(* IEC 61131-3 sources: plcassist-cli/packages/volt-lsp-iec/test-corpus/pro2193/Device/Plc Logic/Application/09 Misc/Library Manager/AlarmManager (part 2) *)

(* ---- ACK_ALARMSTATEMACHINE.fb ---- *)
FUNCTION_BLOCK ACK_ALARMSTATEMACHINE
END_FUNCTION_BLOCK

METHOD DOACKNOWLEDGE : AlarmState
VAR_INPUT
	ECURRENTSTATE : AlarmState;
END_VAR
VAR_OUTPUT
	ESTATETRANSITION : AlarmStateTransition;
END_VAR
END_METHOD

METHOD DOACTIVATE : AlarmState
VAR_INPUT
	ECURRENTSTATE : AlarmState;
END_VAR
END_METHOD

METHOD DODEACTIVATE : AlarmState
VAR_INPUT
	ECURRENTSTATE : AlarmState;
END_VAR
VAR_OUTPUT
	ESTATETRANSITION : AlarmStateTransition;
END_VAR
END_METHOD

(* ---- ACK_ALARMSTATEMACHINE_NOCONFIRM.fb ---- *)
FUNCTION_BLOCK ACK_ALARMSTATEMACHINE_NOCONFIRM EXTENDS Ack_AlarmStateMachine
END_FUNCTION_BLOCK

METHOD DOACKNOWLEDGE : AlarmState
VAR_INPUT
	ECURRENTSTATE : AlarmState;
END_VAR
VAR_OUTPUT
	ESTATETRANSITION : AlarmStateTransition;
END_VAR
END_METHOD

(* ---- ACK_REP_ACK_ALARMSTATEMACHINE.fb ---- *)
FUNCTION_BLOCK ACK_REP_ACK_ALARMSTATEMACHINE
END_FUNCTION_BLOCK

METHOD DOACKNOWLEDGE : AlarmState
VAR_INPUT
	ECURRENTSTATE : AlarmState;
END_VAR
VAR_OUTPUT
	ESTATETRANSITION : AlarmStateTransition;
END_VAR
END_METHOD

METHOD DOACTIVATE : AlarmState
VAR_INPUT
	ECURRENTSTATE : AlarmState;
END_VAR
END_METHOD

METHOD DODEACTIVATE : AlarmState
VAR_INPUT
	ECURRENTSTATE : AlarmState;
END_VAR
VAR_OUTPUT
	ESTATETRANSITION : AlarmStateTransition;
END_VAR
END_METHOD

(* ---- ACK_REP_ACK_ALARMSTATEMACHINE_NOCONFIRM.fb ---- *)
FUNCTION_BLOCK ACK_REP_ACK_ALARMSTATEMACHINE_NOCONFIRM EXTENDS Ack_Rep_Ack_AlarmStateMachine
END_FUNCTION_BLOCK

METHOD DOACKNOWLEDGE : AlarmState
VAR_INPUT
	ECURRENTSTATE : AlarmState;
END_VAR
VAR_OUTPUT
	ESTATETRANSITION : AlarmStateTransition;
END_VAR
END_METHOD

METHOD DODEACTIVATE : AlarmState
VAR_INPUT
	ECURRENTSTATE : AlarmState;
END_VAR
VAR_OUTPUT
	ESTATETRANSITION : AlarmStateTransition;
END_VAR
END_METHOD

(* ---- ACK_REP_ALARMSTATEMACHINE.fb ---- *)
FUNCTION_BLOCK ACK_REP_ALARMSTATEMACHINE
END_FUNCTION_BLOCK

METHOD DOACKNOWLEDGE : AlarmState
VAR_INPUT
	ECURRENTSTATE : AlarmState;
END_VAR
VAR_OUTPUT
	ESTATETRANSITION : AlarmStateTransition;
END_VAR
END_METHOD

METHOD DOACTIVATE : AlarmState
VAR_INPUT
	ECURRENTSTATE : AlarmState;
END_VAR
END_METHOD

METHOD DODEACTIVATE : AlarmState
VAR_INPUT
	ECURRENTSTATE : AlarmState;
END_VAR
VAR_OUTPUT
	ESTATETRANSITION : AlarmStateTransition;
END_VAR
END_METHOD

(* ---- ACK_REP_ALARMSTATEMACHINE_NOCONFIRM.fb ---- *)
FUNCTION_BLOCK ACK_REP_ALARMSTATEMACHINE_NOCONFIRM EXTENDS Ack_Rep_AlarmStateMachine
END_FUNCTION_BLOCK

METHOD DOACKNOWLEDGE : AlarmState
VAR_INPUT
	ECURRENTSTATE : AlarmState;
END_VAR
VAR_OUTPUT
	ESTATETRANSITION : AlarmStateTransition;
END_VAR
END_METHOD

METHOD DODEACTIVATE : AlarmState
VAR_INPUT
	ECURRENTSTATE : AlarmState;
END_VAR
VAR_OUTPUT
	ESTATETRANSITION : AlarmStateTransition;
END_VAR
END_METHOD

(* ---- ACTIVEALARMSTEMPSTORAGE.fb ---- *)
FUNCTION_BLOCK ACTIVEALARMSTEMPSTORAGE
VAR
	_LSTALARMSINFO : COL.IDoubleLinkedList := NULL;
	_LINKEDLISTFACTORY : COL.LinkedListFactory;
	_LISTVALUEELEMFACTORY : ListElementFactory;
END_VAR
END_FUNCTION_BLOCK

METHOD RESTOREALARMS : BOOL
END_METHOD

METHOD STOREALARMS : COL.COLLECTION_ERROR
VAR_INPUT
	PALARMGROUP : IAlarmGroup6;
END_VAR
END_METHOD

METHOD PRVRESTOREADDITIONALALARMINFO : INT
VAR_INPUT
	ITFLISTELEMENT : IListElement;
	PALARMUSED : POINTER TO Alarm;
END_VAR
END_METHOD

METHOD PRVSETALARMINFO : INT
VAR_INPUT
	PALARMSTORED : POINTER TO Alarm;
	PALARMUSED : POINTER TO Alarm;
	ITFLISTELEMENT : IListElement;
END_VAR
END_METHOD

METHOD PRVSTOREACTIVEALARM : BOOL
VAR_INPUT
	ITFLISTELEMENT : IListElement;
	PALARM : POINTER TO Alarm;
END_VAR
END_METHOD

METHOD PRVSTOREALARMS : BOOL
VAR_INPUT
	PALARMGROUP : IAlarmGroup6;
END_VAR
END_METHOD

(* ---- ADAPTERDATABLOCK.fb ---- *)
FUNCTION_BLOCK ADAPTERDATABLOCK
VAR_INPUT
	M_PARRITFALARMSFROMHISTORY : POINTER TO ARRAY [0..0] OF IAlarm2;
	M_PARRALARMSGRPFORHISTORY : POINTER TO ARRAY [0..10] OF POINTER TO AlarmGroupAdapter;
	M_PARRALARMSCLFORHISTORY : POINTER TO ARRAY [0..10] OF POINTER TO AlarmClassAdapter;
	M_ICOUNTALARMSFROMHISTORY : INT;
	M_PAITFALARMCONFIGURATIONS : POINTER TO ARRAY [0..0] OF IAlarmConfiguration;
	M_ICOUNTCONFIGURATIONS : INT;
	M_DITOTALCOUNTROWS : DINT;
END_VAR
VAR
	M_ALARMADAPTER : AlarmAdapter;
	M_ICOUNTROWS : INT;
END_VAR
END_FUNCTION_BLOCK

METHOD GETALARMMETAOBJECTSTUB : IAlarmMetaObjectStub3
VAR_INPUT
	IROW : INT;
	IOFFSET : INT;
END_VAR
END_METHOD

METHOD GETCOUNTROWS : INT
END_METHOD

METHOD HASALARMS : BOOL
END_METHOD

METHOD SETCOUNTROWS : BOOL
VAR_INPUT
	ICOUNT : INT;
END_VAR
END_METHOD

METHOD SETTOTALCOUNTROWS : BOOL
VAR_INPUT
	DICOUNT : DINT;
END_VAR
END_METHOD

(* ---- ALARM.fb ---- *)
FUNCTION_BLOCK ALARM
VAR_INPUT
	M_UIID : ALARM_ID;
	M_UDIID : UDINT;
	M_PALATCHVARIABLES : POINTER TO ARRAY [0..255] OF POINTER TO ValueTypeBundle;
	M_USICOUNTLATCHVARIABLES : USINT;
	M_XDYNVARIABLES : BOOL;
	M_PAPLACEHOLDERINFO : POINTER TO ARRAY [0..255] OF POINTER TO PlaceholderInfo;
	M_USICOUNTMESSAGES : USINT;
END_VAR
VAR
	M_ITFALARMOBSERVATIONTYPE : IAlarmObservationType;
	M_ITFDEACTIVATOR : IDeactivator;
	M_ITFALARMCLASS : IAlarmClass;
	M_ITFALARMGROUP : IAlarmGroup;
	M_ITFALARMGROUPTEMPLATE : IAlarmGroup;
	M_TONDELAYTIME : TIME;
	M_TOFFDELAYTIME : TIME;
	M_LITIMESTAMPACTIVE : Timestamp;
	M_LITIMESTAMPINACTIVE : Timestamp;
	M_LITIMESTAMPACKNOWLEDGE : Timestamp;
	M_LITIMESTAMPLAST : Timestamp;
	M_LITIMESTAMPONDELAY : Timestamp;
	M_LITIMESTAMPOFFDELAY : Timestamp;
	M_IOFFSETACTIVE : INT := -1;
	M_IOFFSETINACTIVE : INT := -1;
	M_IOFFSETACKNOWLEDGE : INT := -1;
	M_IOFFSETLAST : INT := -1;
	M_ESTATE : AlarmState;
	M_XTOACKNOWLEDGE : BOOL;
	M_TIGGERVALUE : ValueTypeBundle;
	M_CURRENTVALUE : ValueTypeBundle;
	M_ITFHIGHERPRIOALARM : IAlarm;
	M_ROWID : CAA.IDENT;
	M_XADDTOLISTOFACTIVEALARMS : BOOL;
	M_XCYCLICUPDATE : BOOL;
	M_XISDEACTIVATEDPREV : BOOL;
	M_SREMDEVICENAME : STRING;
	M_CMTACTIVE : AlarmComment;
	M_CMTACTIVEACK : AlarmComment;
	M_CMTWAITINGCONF : AlarmComment;
	M_CMTNORMAL : AlarmComment;
	M_UDIREALARMREPEATCOUNT : UDINT;
	M_USICOUNTLATCHVARIABLESORIGINAL : INT := -1;
	M_ITFALARM : IAlarm := THIS^;
	ACKNOWLEDGE : BOOL;
	ADDTOLISTOFACTIVEALARMS : BOOL;
	ALARMGROUPTEMPLATE : IAlarmGroup;
	COMMENTACTIVE : POINTER TO WSTRING;
	COMMENTACTIVEACK : POINTER TO WSTRING;
	COMMENTNORMAL : POINTER TO WSTRING;
	COMMENTWAITINGCONF : POINTER TO WSTRING;
	COUNTLATCHVARIABLESORIGINAL : INT;
	CYCLICUPDATE : BOOL;
	ISDEACTIVATEDPREV : BOOL;
	KINDOF : EAlarmType;
	OFFSETACKNOWLEDGE : INT;
	OFFSETACTIVE : INT;
	OFFSETINACTIVE : INT;
	OFFSETLAST : INT;
	REALARMREPEATCOUNT : UDINT;
	REMOTEDEVICENAME : STRING;
	USERIDCOMMENTACTIVE : POINTER TO WSTRING;
	USERIDCOMMENTACTIVEACK : POINTER TO WSTRING;
	USERIDCOMMENTNORMAL : POINTER TO WSTRING;
	USERIDCOMMENTWAITINGCONF : POINTER TO WSTRING;
END_VAR
END_FUNCTION_BLOCK

METHOD ANALYZEPLACEHOLDERS3 : BOOL
VAR_INPUT
	STRINGTYPE : __SYSTEM.TYPE_CLASS;
	IWHICHMESSAGE : INT;
END_VAR
END_METHOD

METHOD FB_EXIT : BOOL
VAR_INPUT
	BINCOPYCODE : BOOL;
END_VAR
END_METHOD

METHOD GETALARMCLASS : IAlarmClass
END_METHOD

METHOD GETALARMGROUP : IAlarmGroup
END_METHOD

METHOD GETHIGHERPRIOALARM : IAlarm
END_METHOD

METHOD GETID : ALARM_ID
END_METHOD

METHOD GETINTERNALID : UDINT
END_METHOD

METHOD GETMESSAGE : CharBufferPtr
VAR_INPUT
	STRINGTYPE : __SYSTEM.TYPE_CLASS;
END_VAR
END_METHOD

METHOD GETOBSERVATIONTYPE : IAlarmObservationType
END_METHOD

METHOD GETROWID : CAA.IDENT
END_METHOD

METHOD GETSTATE : AlarmState
END_METHOD

METHOD ISDEACTIVATED : BOOL
END_METHOD

METHOD SETALARMCLASS
VAR_INPUT
	ITFALARMCLASS : IAlarmClass;
END_VAR
END_METHOD

METHOD SETALARMGROUP
VAR_INPUT
	ITFALARMGROUP : IAlarmGroup;
END_VAR
END_METHOD

METHOD SETHIGHERPRIOALARM
VAR_INPUT
	ITFALARM : IAlarm;
END_VAR
END_METHOD

METHOD SETOBSERVATIONTYPE
VAR_INPUT
	ITFOBSERVATIONTYPE : IAlarmObservationType;
END_VAR
END_METHOD

METHOD SETROWID
VAR_INPUT
	ROWID : CAA.IDENT;
END_VAR
END_METHOD

METHOD SETTIMESTAMP
VAR_INPUT
	LICURRTIMESTAMP : Timestamp;
	ESTATE : AlarmState;
	ESTATETRANSITION : AlarmStateTransition;
END_VAR
END_METHOD

METHOD SETALARMSTATE
VAR_INPUT
	EALARMSTATE : AlarmState;
END_VAR
END_METHOD

METHOD SETCURRENTVALUE
VAR_INPUT
	ITFTYPEDVALUECURRENT : ITypedValue;
END_VAR
END_METHOD

METHOD SETID
VAR_INPUT
	UIID : ALARM_ID;
END_VAR
END_METHOD

METHOD SETINTERNALID
VAR_INPUT
	UDIID : UDINT;
END_VAR
END_METHOD

METHOD SETLATCHVAR1VALUE
VAR_INPUT
	ITFTYPEDVALUELATCHVAR1 : ITypedValue;
END_VAR
END_METHOD

METHOD SETLATCHVAR2VALUE
VAR_INPUT
	ITFTYPEDVALUELATCHVAR2 : ITypedValue;
END_VAR
END_METHOD

METHOD SETTIMESTAMPACKNOWLEDGE
VAR_INPUT
	LITIMESTAMPACKNOWLEDGE : Timestamp;
END_VAR
END_METHOD

METHOD SETTIMESTAMPACTIVE
VAR_INPUT
	LITIMESTAMPACTIVE : Timestamp;
END_VAR
END_METHOD

METHOD SETTIMESTAMPINACTIVE
VAR_INPUT
	LITIMESTAMPINACTIVE : Timestamp;
END_VAR
END_METHOD

METHOD SETTIMESTAMPLAST
VAR_INPUT
	LITIMESTAMPLAST : Timestamp;
END_VAR
END_METHOD

METHOD SETTRIGGERVALUE
VAR_INPUT
	ITFTYPEDVALUETRIGGER : ITypedValue;
END_VAR
END_METHOD

METHOD GETCOUNTLATCHVARIABLES : USINT
END_METHOD

METHOD GETCOUNTMESSAGES : USINT
END_METHOD

METHOD GETLATCHVARVALUE : ITypedValue
VAR_INPUT
	IWHICHLATCHVAR : INT;
END_VAR
END_METHOD

METHOD GETMESSAGE2 : CharBufferPtr
VAR_INPUT
	STRINGTYPE : __SYSTEM.TYPE_CLASS;
	IWHICHMESSAGE : INT;
END_VAR
END_METHOD

METHOD SETLATCHVARVALUE
VAR_INPUT
	IWHICHLATCHVAR : INT;
	ITFTYPEDVALUELATCHVAR : ITypedValue;
END_VAR
END_METHOD

METHOD SETTIMESTAMP2
VAR_INPUT
	LICURRTIMESTAMP : Timestamp;
	IOFFSET : INT;
	ESTATE : AlarmState;
	ESTATETRANSITION : AlarmStateTransition;
END_VAR
END_METHOD

METHOD GETLATCHVARIABLESADDRESS
VAR_OUTPUT
	PALATCHVARIABLES : POINTER TO BYTE;
	USICOUNTLATCHVARIABLES : USINT;
END_VAR
END_METHOD

METHOD SETLATCHVARIABLESADDRESS
VAR_INPUT
	PALATCHVARIABLES : POINTER TO BYTE;
	USICOUNTLATCHVARIABLES : USINT;
END_VAR
END_METHOD

METHOD ANALYZEPLACEHOLDERS
VAR_INPUT
	STRINGTYPE : __SYSTEM.TYPE_CLASS;
END_VAR
END_METHOD

METHOD GETCOUNTPLACEHOLDERS : SINT
END_METHOD

METHOD GETPLACEHOLDER : PlaceholderOccurrence
VAR_INPUT
	SIWHICHPLACEHOLDER : SINT;
END_VAR
END_METHOD

METHOD HASPLACEHOLDERREQUIRINGCYCLICALLYUPDATE : BOOL
END_METHOD

METHOD HASPLACEHOLDERS : BOOL
END_METHOD

METHOD ISOPTIMIZEDPLACEHOLDERREPLACEMENTSUPPORTED : BOOL
END_METHOD

METHOD ANALYZEPLACEHOLDERS2
VAR_INPUT
	STRINGTYPE : __SYSTEM.TYPE_CLASS;
	IWHICHMESSAGE : INT;
END_VAR
END_METHOD

METHOD GETCOUNTPLACEHOLDERS2 : SINT
VAR_INPUT
	IWHICHMESSAGE : INT;
END_VAR
END_METHOD

METHOD GETPLACEHOLDER2 : PlaceholderOccurrence
VAR_INPUT
	SIWHICHPLACEHOLDER : SINT;
	IWHICHMESSAGE : INT;
END_VAR
END_METHOD

METHOD HASPLACEHOLDERREQUIRINGCYCLICALLYUPDATE2 : BOOL
VAR_INPUT
	IWHICHMESSAGE : INT;
END_VAR
END_METHOD

METHOD HASPLACEHOLDERS2 : BOOL
VAR_INPUT
	IWHICHMESSAGE : INT;
END_VAR
END_METHOD

METHOD ISOPTIMIZEDPLACEHOLDERREPLACEMENTSUPPORTED2 : BOOL
VAR_INPUT
	IWHICHMESSAGE : INT;
END_VAR
END_METHOD

METHOD CANBEACTIVATED : BOOL
END_METHOD

METHOD CANBEDEACTIVATED : BOOL
END_METHOD

METHOD DETERMINETIMESTAMP
VAR_INPUT
	ESTATE : AlarmState;
	ESTATETRANSITION : AlarmStateTransition;
END_VAR
END_METHOD

METHOD GETALARM : IAlarm
END_METHOD

METHOD GETLATCHVARIABLESADDRESSDIRECT : BOOL
VAR_OUTPUT
	PALATCHVARIABLES : POINTER TO BYTE;
	USICOUNTLATCHVARIABLES : USINT;
END_VAR
END_METHOD

METHOD HANDLEAUTORESETDIGITALALARMS : BOOL
END_METHOD

METHOD INVALIDATEMESSAGEFLAGS
END_METHOD

METHOD RETRIEVECURRENTVALUE
VAR_INPUT
	ITFVALUEPROVIDER : IValueProvider;
END_VAR
END_METHOD

METHOD RETRIEVELATCHVARVALUE
VAR_INPUT
	IWHICHLATCHVARIABLE : INT;
	ITFVALUEPROVIDER : IValueProvider;
END_VAR
END_METHOD

METHOD RETRIEVELATCHVARVALUES
VAR_INPUT
	ITFVALUEPROVIDER : IValueProvider;
END_VAR
END_METHOD

METHOD RETRIEVETRIGGERVALUE
VAR_INPUT
	ITFVALUEPROVIDER : IValueProvider;
END_VAR
END_METHOD

METHOD SETACKNOWLEDGE : BOOL
VAR_INPUT
	PWSCOMMENT : POINTER TO WSTRING;
	PWSUSERID : POINTER TO WSTRING;
END_VAR
END_METHOD

METHOD SETACKNOWLEDGELOCKED : BOOL
VAR_INPUT
	PWSCOMMENT : POINTER TO WSTRING;
	PWSUSERID : POINTER TO WSTRING;
END_VAR
END_METHOD

METHOD SETCOMMENT : UDINT
VAR_INPUT
	PWSCOMMENT : POINTER TO WSTRING;
	PWSUSERID : POINTER TO WSTRING;
END_VAR
END_METHOD

METHOD SETCOMMENTDIRECTLY
VAR_INPUT
	PALARMOTHER : POINTER TO Alarm;
END_VAR
END_METHOD

METHOD SETDEACTIVATOR
VAR_INPUT
	ITFDEACTIVATOR : IDeactivator;
END_VAR
END_METHOD

METHOD SETOFFDELAYTIME
VAR_INPUT
	TTIME : TIME;
END_VAR
END_METHOD

METHOD SETONDELAYTIME
VAR_INPUT
	TTIME : TIME;
END_VAR
END_METHOD

METHOD SETREALARMREPEATCOUNTDIRECTLY
VAR_INPUT
	UDIREALARMREPEATCOUNT : UDINT;
END_VAR
END_METHOD

METHOD SETSTATE
VAR_INPUT
	ESTATE : AlarmState;
	ESTATETRANSITION : AlarmStateTransition;
END_VAR
END_METHOD

METHOD SETTIMESTAMPOFFDELAY
VAR_INPUT
	XRESET : BOOL;
END_VAR
END_METHOD

METHOD SETTIMESTAMPDELAY
VAR_INPUT
	XRESET : BOOL;
	TDELAY : TIME;
END_VAR
VAR_IN_OUT
	LITIMESTAMPDELAY : Timestamp;
END_VAR
END_METHOD

METHOD SETTIMESTAMPOFFDELAYDIRECTLY
VAR_INPUT
	LITIMESTAMPOFFDELAY : Timestamp;
END_VAR
END_METHOD

METHOD SETTIMESTAMPONDELAY
VAR_INPUT
	XRESET : BOOL;
END_VAR
END_METHOD

METHOD SETTIMESTAMPONDELAYDIRECTLY
VAR_INPUT
	LITIMESTAMPONDELAY : Timestamp;
END_VAR
END_METHOD

METHOD SETTRIGGERVALUEDIRECTLY
VAR_INPUT
	TRIGGERVALUE : ValueTypeBundle;
END_VAR
END_METHOD

METHOD ISCOMMENTTOSTATENORMAL : BOOL
END_METHOD

METHOD RESETALARMCOMMENTS
END_METHOD

METHOD RESETFORNEWCYCLE
END_METHOD

METHOD PRVCHECKPOSTALARM
VAR_INPUT
	ESTATE : AlarmState;
	EOLDSTATE : AlarmState;
	XFORCEUPDATE : BOOL;
END_VAR
END_METHOD

METHOD PRVCOPYFROMTYPEDVALUE
VAR_INPUT
	PVALUETYPEBUNDLETARGET : POINTER TO ValueTypeBundle;
	ITFTYPEDVALUESOURCE : ITypedValue;
END_VAR
END_METHOD

METHOD GETTIMESTAMPACKNOWLEDGE : Timestamp
END_METHOD

METHOD GETTIMESTAMPACTIVE : Timestamp
END_METHOD

METHOD GETTIMESTAMPINACTIVE : Timestamp
END_METHOD

METHOD GETTIMESTAMPLAST : Timestamp
END_METHOD

METHOD GETCURRENTVALUE : ITypedValue
END_METHOD

METHOD GETLATCHVAR1VALUE : ITypedValue
END_METHOD

METHOD GETLATCHVAR2VALUE : ITypedValue
END_METHOD

METHOD GETTRIGGERVALUE : ITypedValue
END_METHOD

(* ---- ALARMADAPTER.fb ---- *)
FUNCTION_BLOCK ALARMADAPTER
VAR_INPUT
	M_ITFALARM2 : IAlarm2;
	M_PALARMGROUP : POINTER TO AlarmGroupAdapter;
	M_PALARMCLASS : POINTER TO AlarmClassAdapter;
	M_PAITFALARMCONFIGURATIONS : POINTER TO ARRAY [0..0] OF IAlarmConfiguration;
	M_ICOUNTCONFIGURATIONS : INT;
END_VAR
VAR
	M_PLIVALUE : POINTER TO LINT;
	ALARMCLASSINTERNALID : UDINT;
	ALARMGROUPINTERNALID : UDINT;
	ALARMINTERNALID : UDINT;
	OFFSETACKNOWLEDGE : INT;
	OFFSETACTIVE : INT;
	OFFSETINACTIVE : INT;
	OFFSETLAST : INT;
	PROXYNAME : STRING;
	REMOTEALARMCLASSNAME : STRING;
	REMOTEALARMGROUPNAME : STRING;
	REMOTEALARMSTRINGID : STRING;
	REMOTEALARMTEXTLIST : STRING;
END_VAR
END_FUNCTION_BLOCK

METHOD INITIALIZE
END_METHOD

METHOD SETALARM
VAR_INPUT
	PALARM : POINTER TO Alarm;
END_VAR
END_METHOD

METHOD SETALARMGROUP
VAR_INPUT
	SALARMGROUP : STRING;
END_VAR
END_METHOD

METHOD SETCURRENTVALUE
VAR_INPUT
	ITFTYPEDVALUECURRENT : AlarmManager_Interfaces.ITypedValue;
END_VAR
END_METHOD

METHOD SETID
VAR_INPUT
	UIID : ALARM_ID;
END_VAR
END_METHOD

METHOD SETLATCHVAR1VALUE
VAR_INPUT
	ITFTYPEDVALUELATCHVAR1 : AlarmManager_Interfaces.ITypedValue;
END_VAR
END_METHOD

METHOD SETLATCHVAR2VALUE
VAR_INPUT
	ITFTYPEDVALUELATCHVAR2 : AlarmManager_Interfaces.ITypedValue;
END_VAR
END_METHOD

METHOD SETSTATE
VAR_INPUT
	ISTATE : INT;
END_VAR
END_METHOD

METHOD SETTIMESTAMPACKNOWLEDGE
VAR_INPUT
	LITIMESTAMPACKNOWLEDGE : Timestamp;
END_VAR
END_METHOD

METHOD SETTIMESTAMPACTIVE
VAR_INPUT
	LITIMESTAMPACTIVE : Timestamp;
END_VAR
END_METHOD

METHOD SETTIMESTAMPINACTIVE
VAR_INPUT
	LITIMESTAMPINACTIVE : Timestamp;
END_VAR
END_METHOD

METHOD SETTIMESTAMPLAST
VAR_INPUT
	LITIMESTAMPLAST : Timestamp;
END_VAR
END_METHOD

METHOD SETTRIGGERVALUE
VAR_INPUT
	ITFTYPEDVALUETRIGGER : AlarmManager_Interfaces.ITypedValue;
END_VAR
END_METHOD

METHOD GETPRIORITY : BYTE
END_METHOD

METHOD SETPRIORITY
VAR_INPUT
	BYPRIORITY : BYTE;
END_VAR
END_METHOD

METHOD GETCOUNTLATCHVARIABLES : USINT
END_METHOD

METHOD SETLATCHVARVALUE
VAR_INPUT
	IWHICHLATCHVAR : INT;
	ITFTYPEDVALUELATCHVAR : ITypedValue;
END_VAR
END_METHOD

METHOD PRVPREPARELATCHVARVALUE : ValueTypeBundle
VAR_INPUT
	ITFTYPEDVALUELATCHVAR : AlarmManager_Interfaces.ITypedValue;
END_VAR
END_METHOD

METHOD GETALARM : POINTER TO Alarm
END_METHOD

METHOD GETALARMGROUP : STRING
END_METHOD

METHOD GETCHECKSUM : UDINT
END_METHOD

METHOD GETCURRENTVALUE : AlarmManager_Interfaces.ITypedValue
END_METHOD

METHOD GETID : ALARM_ID
END_METHOD

METHOD GETLATCHVAR1VALUE : AlarmManager_Interfaces.ITypedValue
END_METHOD

METHOD GETLATCHVAR2VALUE : AlarmManager_Interfaces.ITypedValue
END_METHOD

METHOD GETSTATE : INT
END_METHOD

METHOD GETTIMESTAMPACKNOWLEDGE : Timestamp
END_METHOD

METHOD GETTIMESTAMPACTIVE : Timestamp
END_METHOD

METHOD GETTIMESTAMPINACTIVE : Timestamp
END_METHOD

METHOD GETTIMESTAMPLAST : Timestamp
END_METHOD

METHOD GETTRIGGERVALUE : AlarmManager_Interfaces.ITypedValue
END_METHOD

METHOD SETACKNOWLEDGE
VAR_INPUT
	BACKNOWLEDGEMULTIPLE : BOOL;
END_VAR
END_METHOD

METHOD SWAPVALUES
END_METHOD

METHOD GETACKNOWLEDGE : BOOL
END_METHOD

METHOD GETACKNOWLEDGEMULTIPLE : BOOL
END_METHOD

METHOD GETALARMCLASS : STRING
END_METHOD

METHOD GETSTRINGID : STRING
END_METHOD

METHOD GETTESTLISTNAME : STRING
END_METHOD

METHOD RESETACKNOWLEDGE
END_METHOD

METHOD SETALARMCLASS
VAR_INPUT
	SALARMCLASS : STRING;
END_VAR
END_METHOD

METHOD SETSTRINGID
VAR_INPUT
	SID : STRING;
END_VAR
END_METHOD

METHOD SETTESTLISTNAME
VAR_INPUT
	STESTLISTNAME : STRING;
END_VAR
END_METHOD

METHOD SETACKNOWLEDGE2
VAR_INPUT
	BACKNOWLEDGEMULTIPLE : BOOL;
END_VAR
END_METHOD

METHOD GETLATCHVARVALUE : ITypedValue2
VAR_INPUT
	IWHICHLATCHVAR : INT;
END_VAR
END_METHOD

(* ---- ALARMAPIOBSERVATIONTYPE.fb ---- *)
FUNCTION_BLOCK ALARMAPIOBSERVATIONTYPE
VAR
	M_XISACTIVE : BOOL;
	ALARMCONDITIONACTIVE : BOOL;
END_VAR
END_FUNCTION_BLOCK

METHOD ISACTIVE : BOOL
VAR_INPUT
	ECURRSTATE : AlarmState;
END_VAR
END_METHOD

METHOD ISIMMEDIATELYACTIVE : BOOL
END_METHOD

(* ---- ALARMCLASS.fb ---- *)
FUNCTION_BLOCK ALARMCLASS
VAR
	M_UDIID : UDINT;
	M_USIPRIORITY : USINT;
	M_XARCHIVING : BOOL;
	M_EACKNOWLEDGEMETHOD : AcknowledgeMethod;
	M_XACKNOWLEDGESEPARATELY : BOOL;
	M_XAUTORESETDIGITALALARMS : BOOL;
	M_XACKINSTEADOFCONFIRM : BOOL;
	M_PAITFALARMNOTIFIABLES : POINTER TO ARRAY [0..0] OF IAlarmNotifiable;
	M_ICOUNTNOTIFIABLES : INT;
	M_SNAME : STRING;
	M_PAPDISPLAYOPTIONS : POINTER TO ARRAY [AlarmState.Normal..AlarmState.ActiveAcknowledged] OF POINTER TO DisplayOptions;
	M_TREALARMTIME : TIME;
	REALARMTIME : TIME;
END_VAR
END_FUNCTION_BLOCK

METHOD SETACKINSTEADOFCONFIRM : BOOL
VAR_INPUT
	XACKINSTEADOFCONFIRM : BOOL;
END_VAR
END_METHOD

METHOD SETACKNOWLEDGEMETHOD
VAR_INPUT
	EACKNOWLEDGEMETHOD : AcknowledgeMethod;
END_VAR
END_METHOD

METHOD SETACKNOWLEDGESEPARATELY
VAR_INPUT
	XACKNOWLEDGESEPARATELY : BOOL;
END_VAR
END_METHOD

METHOD SETALARMNOTIFIABLES
END_METHOD

METHOD SETARCHIVING
VAR_INPUT
	XARCHIVING : BOOL;
END_VAR
END_METHOD

METHOD SETAUTORESETDIGITALALARMS
VAR_INPUT
	XAUTORESETDIGITALALARMS : BOOL;
END_VAR
END_METHOD

METHOD SETDISPLAYOPTIONS
END_METHOD

METHOD SETINTERNALID
VAR_INPUT
	UDIID : UDINT;
END_VAR
END_METHOD

METHOD SETNAME
VAR_INPUT
	SNAME : STRING;
END_VAR
END_METHOD

METHOD SETPRIORITY
VAR_INPUT
	USIPRIORITY : USINT;
END_VAR
END_METHOD

METHOD SETREALARMTIME
VAR_INPUT
	T : TIME;
END_VAR
END_METHOD

METHOD GETACKNOWLEDGEMETHOD : AcknowledgeMethod
END_METHOD

METHOD GETALARMSTATEMACHINE : IAlarmStateMachine
END_METHOD

METHOD GETDISPLAYOPTIONS : POINTER TO DisplayOptions
VAR_INPUT
	ESTATE : AlarmState;
END_VAR
END_METHOD

METHOD GETINTERNALID : UDINT
END_METHOD

METHOD GETNAME : STRING
END_METHOD

METHOD GETPRIORITY : USINT
END_METHOD

METHOD ISACKNOWLEDGESEPARATELY : BOOL
END_METHOD

METHOD ACKINSTEADOFCONFIRM : BOOL
END_METHOD

METHOD AUTORESETDIGITALALARMS : BOOL
END_METHOD

METHOD GETALARMCLASSOBJECTCHECKSUM : LINT
END_METHOD

METHOD GETARCHIVING : BOOL
END_METHOD

METHOD NOTIFYNOTIFIABLES
VAR_INPUT
	ESTATETRANSITION : AlarmStateTransition;
	ITFALARM : IAlarm;
END_VAR
END_METHOD

(* ---- ALARMCLASSADAPTER.fb ---- *)
FUNCTION_BLOCK ALARMCLASSADAPTER EXTENDS AlarmClassContainerBase
END_FUNCTION_BLOCK

(* ---- ALARMCLASSCOMPARER.fb ---- *)
FUNCTION_BLOCK ALARMCLASSCOMPARER EXTENDS TSLastComparer
END_FUNCTION_BLOCK

METHOD COMPARE : INT
VAR_INPUT
	DIINDEXALARM1 : DINT;
	DIINDEXALARM2 : DINT;
END_VAR
END_METHOD

(* ---- ALARMCLASSCONTAINERBASE.fb ---- *)
FUNCTION_BLOCK ALARMCLASSCONTAINERBASE
VAR_INPUT
	M_UDIID : UDINT;
	M_SNAME : STRING;
	M_USIPRIORITY : USINT;
	M_ADISPLAYOPTIONS : ARRAY [AlarmState.Normal..AlarmState.ActiveAcknowledged] OF DisplayOptions;
END_VAR
END_FUNCTION_BLOCK

METHOD GETDISPLAYOPTIONS : POINTER TO DisplayOptions
VAR_INPUT
	ESTATE : AlarmState;
END_VAR
END_METHOD

METHOD GETINTERNALID : UDINT
END_METHOD

METHOD GETNAME : STRING
END_METHOD

METHOD GETPRIORITY : USINT
END_METHOD

METHOD GETACKNOWLEDGEMETHOD : AcknowledgeMethod
END_METHOD

METHOD GETALARMSTATEMACHINE : IAlarmStateMachine
END_METHOD

METHOD ISACKNOWLEDGESEPARATELY : BOOL
END_METHOD

(* ---- ALARMCLASSMOCK.fb ---- *)
FUNCTION_BLOCK ALARMCLASSMOCK EXTENDS AlarmClassContainerBase
END_FUNCTION_BLOCK

METHOD SETVALUES
VAR_INPUT
	ISET : INT;
END_VAR
END_METHOD

(* ---- ALARMCOMMENTHELPER.fb ---- *)
FUNCTION_BLOCK ALARMCOMMENTHELPER
END_FUNCTION_BLOCK

METHOD COPYWSTRINGTOALARMCOMMENT : BOOL
VAR_INPUT
	PWSCOMMENT : POINTER TO WSTRING;
	PWSUSERID : POINTER TO WSTRING;
END_VAR
VAR_IN_OUT
	ALARMCOMMENT : AlarmComment;
END_VAR
END_METHOD

METHOD FREEALARMCOMMENT : BOOL
VAR_IN_OUT
	ALARMCOMMENT : AlarmComment;
END_VAR
END_METHOD

(* ---- ALARMCONTAINER.fb ---- *)
FUNCTION_BLOCK ALARMCONTAINER EXTENDS AlarmContainerBase
VAR_INPUT
	M_ALARMGROUP : AlarmGroupContainerBase;
	M_ALARMCLASS : AlarmClassContainerBase;
	M_STEXTLISTINDEX : STRING;
	M_PALATCHVARIABLES : POINTER TO ARRAY [0..255] OF POINTER TO ValueTypeBundle;
	M_SPROXYNAME : STRING;
	M_IFTPROXY : IProxy;
END_VAR
VAR
	REMOTEDEVICENAME : STRING;
END_VAR
END_FUNCTION_BLOCK

METHOD FB_EXIT : BOOL
VAR_INPUT
	BINCOPYCODE : BOOL;
END_VAR
END_METHOD

METHOD FB_INIT : BOOL
VAR_INPUT
	BINITRETAINS : BOOL;
	BINCOPYCODE : BOOL;
END_VAR
END_METHOD

METHOD PRVCOPYFROMTYPEDVALUE
VAR_INPUT
	PVALUETYPEBUNDLETARGET : POINTER TO ValueTypeBundle;
	ITFTYPEDVALUESOURCE : ITypedValue;
END_VAR
END_METHOD

METHOD GETCURRENTVALUE : ITypedValue
END_METHOD

METHOD GETLATCHVAR1VALUE : ITypedValue
END_METHOD

METHOD GETLATCHVAR2VALUE : ITypedValue
END_METHOD

METHOD GETLATCHVARVALUE : ITypedValue
VAR_INPUT
	IWHICHLATCHVAR : INT;
END_VAR
END_METHOD

METHOD GETMESSAGE : Stu.CharBufferPtr
VAR_INPUT
	STRINGTYPE : __SYSTEM.TYPE_CLASS;
END_VAR
END_METHOD

METHOD GETMESSAGE2 : Stu.CharBufferPtr
VAR_INPUT
	STRINGTYPE : __SYSTEM.TYPE_CLASS;
	IWHICHMESSAGE : INT;
END_VAR
END_METHOD

METHOD GETTRIGGERVALUE : ITypedValue
END_METHOD

METHOD SETCURRENTVALUE
VAR_INPUT
	ITFTYPEDVALUECURRENT : ITypedValue;
END_VAR
END_METHOD

METHOD SETLATCHVARVALUE
VAR_INPUT
	IWHICHLATCHVAR : INT;
	ITFTYPEDVALUELATCHVAR : ITypedValue;
END_VAR
END_METHOD

METHOD SETTRIGGERVALUE
VAR_INPUT
	ITFTYPEDVALUETRIGGER : ITypedValue;
END_VAR
END_METHOD

(* ---- ALARMCONTAINERBASE.fb ---- *)
FUNCTION_BLOCK ALARMCONTAINERBASE
VAR_INPUT
	M_ITFALARMGROUP : IAlarmGroup;
	M_ITFALARMCLASS : IAlarmClass;
	M_TIGGERVALUE : ValueTypeBundle;
	M_ITIGGERVALUE : INT;
	M_CURRENTVALUE : ValueTypeBundle;
	M_ICURRENTVALUE : INT;
	M_LATCHVARIABLE1 : ValueTypeBundle;
	M_LATCHVARIABLE2 : ValueTypeBundle;
	M_LATCHVARIABLE3 : ValueTypeBundle;
	M_SVALUE : STRING;
	M_WSVALUE : WSTRING;
	M_USICOUNTLATCHVARIABLES : USINT;
	M_USICOUNTMESSAGES : USINT;
	M_UIID : ALARM_ID;
	M_UDIID : UDINT;
	M_ESTATE : AlarmState;
	M_LITIMESTAMPACKNOWLEDGE : Timestamp;
	M_LITIMESTAMPACTIVE : Timestamp;
	M_LITIMESTAMPINACTIVE : Timestamp;
	M_LITIMESTAMPLAST : Timestamp;
	M_IOFFSETACTIVE : INT;
	M_IOFFSETINACTIVE : INT;
	M_IOFFSETACKNOWLEDGE : INT;
	M_IOFFSETLAST : INT;
END_VAR
VAR
	ADDTOLISTOFACTIVEALARMS : BOOL;
	KINDOF : EAlarmType;
	OFFSETACKNOWLEDGE : INT;
	OFFSETACTIVE : INT;
	OFFSETINACTIVE : INT;
	OFFSETLAST : INT;
END_VAR
END_FUNCTION_BLOCK

METHOD GETALARMCLASS : IAlarmClass
END_METHOD

METHOD GETALARMGROUP : IAlarmGroup
END_METHOD

METHOD GETCOUNTLATCHVARIABLES : USINT
END_METHOD

METHOD GETCOUNTMESSAGES : USINT
END_METHOD

METHOD GETID : ALARM_ID
END_METHOD

METHOD GETINTERNALID : UDINT
END_METHOD

METHOD GETSTATE : AlarmState
END_METHOD

METHOD GETTIMESTAMPACKNOWLEDGE : Timestamp
END_METHOD

METHOD GETTIMESTAMPACTIVE : Timestamp
END_METHOD

METHOD GETTIMESTAMPINACTIVE : Timestamp
END_METHOD

METHOD GETTIMESTAMPLAST : Timestamp
END_METHOD

METHOD ANALYZEPLACEHOLDERS
VAR_INPUT
	STRINGTYPE : __SYSTEM.TYPE_CLASS;
END_VAR
END_METHOD

METHOD ANALYZEPLACEHOLDERS2
VAR_INPUT
	STRINGTYPE : __SYSTEM.TYPE_CLASS;
	IWHICHMESSAGE : INT;
END_VAR
END_METHOD

METHOD GETCOUNTPLACEHOLDERS : SINT
END_METHOD

METHOD GETCOUNTPLACEHOLDERS2 : SINT
VAR_INPUT
	IWHICHMESSAGE : INT;
END_VAR
END_METHOD

METHOD GETCURRENTVALUE : AlarmManager_Interfaces.ITypedValue
END_METHOD

METHOD GETLATCHVAR1VALUE : AlarmManager_Interfaces.ITypedValue
END_METHOD

METHOD GETLATCHVAR2VALUE : AlarmManager_Interfaces.ITypedValue
END_METHOD

METHOD GETLATCHVARVALUE : ITypedValue
VAR_INPUT
	IWHICHLATCHVAR : INT;
END_VAR
END_METHOD

METHOD GETMESSAGE : Stu.CharBufferPtr
VAR_INPUT
	STRINGTYPE : __SYSTEM.TYPE_CLASS;
END_VAR
END_METHOD

METHOD GETMESSAGE2 : Stu.CharBufferPtr
VAR_INPUT
	STRINGTYPE : __SYSTEM.TYPE_CLASS;
	IWHICHMESSAGE : INT;
END_VAR
END_METHOD

METHOD GETOBSERVATIONTYPE : IAlarmObservationType
END_METHOD

METHOD GETPLACEHOLDER : PlaceholderOccurrence
VAR_INPUT
	SIWHICHPLACEHOLDER : SINT;
END_VAR
END_METHOD

METHOD GETPLACEHOLDER2 : PlaceholderOccurrence
VAR_INPUT
	SIWHICHPLACEHOLDER : SINT;
	IWHICHMESSAGE : INT;
END_VAR
END_METHOD

METHOD GETROWID : CAA.IDENT
END_METHOD

METHOD GETTRIGGERVALUE : AlarmManager_Interfaces.ITypedValue
END_METHOD

METHOD HASPLACEHOLDERREQUIRINGCYCLICALLYUPDATE : BOOL
END_METHOD

METHOD HASPLACEHOLDERREQUIRINGCYCLICALLYUPDATE2 : BOOL
VAR_INPUT
	IWHICHMESSAGE : INT;
END_VAR
END_METHOD

METHOD HASPLACEHOLDERS : BOOL
END_METHOD

METHOD HASPLACEHOLDERS2 : BOOL
VAR_INPUT
	IWHICHMESSAGE : INT;
END_VAR
END_METHOD

METHOD ISDEACTIVATED : BOOL
END_METHOD

METHOD ISOPTIMIZEDPLACEHOLDERREPLACEMENTSUPPORTED : BOOL
END_METHOD

METHOD ISOPTIMIZEDPLACEHOLDERREPLACEMENTSUPPORTED2 : BOOL
VAR_INPUT
	IWHICHMESSAGE : INT;
END_VAR
END_METHOD

METHOD SETALARMCLASS
VAR_INPUT
	ITFALARMCLASS : IAlarmClass;
END_VAR
END_METHOD

METHOD SETALARMGROUP
VAR_INPUT
	ITFALARMGROUP : IAlarmGroup;
END_VAR
END_METHOD

METHOD SETALARMSTATE
VAR_INPUT
	EALARMSTATE : AlarmState;
END_VAR
END_METHOD

METHOD SETCURRENTVALUE
VAR_INPUT
	ITFTYPEDVALUECURRENT : ITypedValue;
END_VAR
END_METHOD

METHOD SETHIGHERPRIOALARM
VAR_INPUT
	ITFALARM : IAlarm;
END_VAR
END_METHOD

METHOD SETLATCHVAR1VALUE
VAR_INPUT
	ITFTYPEDVALUELATCHVAR1 : ITypedValue;
END_VAR
END_METHOD

METHOD SETLATCHVAR2VALUE
VAR_INPUT
	ITFTYPEDVALUELATCHVAR2 : ITypedValue;
END_VAR
END_METHOD

METHOD SETLATCHVARVALUE
VAR_INPUT
	IWHICHLATCHVAR : INT;
	ITFTYPEDVALUELATCHVAR : ITypedValue;
END_VAR
END_METHOD

METHOD SETOBSERVATIONTYPE
VAR_INPUT
	ITFOBSERVATIONTYPE : IAlarmObservationType;
END_VAR
END_METHOD

METHOD SETROWID
VAR_INPUT
	ROWID : CAA.IDENT;
END_VAR
END_METHOD

METHOD SETTIMESTAMP
VAR_INPUT
	LICURRTIMESTAMP : Timestamp;
	ESTATE : AlarmState;
	ESTATETRANSITION : AlarmStateTransition;
END_VAR
END_METHOD

METHOD SETTIMESTAMP2
VAR_INPUT
	LICURRTIMESTAMP : Timestamp;
	IOFFSET : INT;
	ESTATE : AlarmState;
	ESTATETRANSITION : AlarmStateTransition;
END_VAR
END_METHOD

METHOD SETTRIGGERVALUE
VAR_INPUT
	ITFTYPEDVALUETRIGGER : ITypedValue;
END_VAR
END_METHOD

METHOD SETID
VAR_INPUT
	UIID : ALARM_ID;
END_VAR
END_METHOD

METHOD SETINTERNALID
VAR_INPUT
	UDIID : UDINT;
END_VAR
END_METHOD

METHOD SETTIMESTAMPACKNOWLEDGE
VAR_INPUT
	LITIMESTAMPACKNOWLEDGE : Timestamp;
END_VAR
END_METHOD

METHOD SETTIMESTAMPACTIVE
VAR_INPUT
	LITIMESTAMPACTIVE : Timestamp;
END_VAR
END_METHOD

METHOD SETTIMESTAMPINACTIVE
VAR_INPUT
	LITIMESTAMPINACTIVE : Timestamp;
END_VAR
END_METHOD

METHOD SETTIMESTAMPLAST
VAR_INPUT
	LITIMESTAMPLAST : Timestamp;
END_VAR
END_METHOD

(* ---- ALARMEVALUATOR.fb ---- *)
FUNCTION_BLOCK ALARMEVALUATOR
END_FUNCTION_BLOCK

METHOD CHECKDEACTIVATION : AlarmState
VAR_INPUT
	ECURRSTATE : AlarmState;
	ITFALARMSTATEMACHINE : IAlarmStateMachine;
END_VAR
VAR_IN_OUT
	ALARM : Alarm;
	ESTATETRANSITION : AlarmStateTransition;
END_VAR
END_METHOD

METHOD CHECKREACTIVATION : AlarmState
VAR_INPUT
	ECURRSTATE : AlarmState;
	ITFALARMSTATEMACHINE : IAlarmStateMachine;
END_VAR
VAR_OUTPUT
	ESTATETRANSITION : AlarmStateTransition;
END_VAR
VAR_IN_OUT
	ALARM : Alarm;
END_VAR
END_METHOD

METHOD ISREALARMING : BOOL
VAR_IN_OUT
	ALARM : Alarm;
END_VAR
END_METHOD

METHOD PREPROCESSALARMACTIVATION
VAR_INPUT
	ALARM : REFERENCE TO Alarm;
	ITFVALUEPROVIDER : IValueProvider;
END_VAR
END_METHOD

METHOD PRVPREPROCESSEVENTACTIVATION
VAR_INPUT
	EVENT : REFERENCE TO Alarm;
END_VAR
VAR_OUTPUT
	BEVENTNEEDEDSTORAGELIMITCOUNT : BOOL;
END_VAR
END_METHOD

METHOD PRVPROCESSACKNOWLEDGEMENT
VAR_INPUT
	ALARM : REFERENCE TO Alarm;
END_VAR
END_METHOD

METHOD PRVPROCESSHIGHERPRIORITYALARM
VAR_INPUT
	ALARM : REFERENCE TO Alarm;
END_VAR
END_METHOD

(* ---- ALARMGROUP.fb ---- *)
FUNCTION_BLOCK ALARMGROUP
VAR_INPUT
	M_ITFALARMSTORAGE : IDatabaseFileAlarmStorage;
	M_SNAME : STRING;
END_VAR
VAR
	M_PAPALARMS : POINTER TO ARRAY [0..0] OF POINTER TO Alarm;
	M_ICOUNTALARMS : INT;
	M_USIALARMGROUPID : ALARMGROUP_ID;
	_ALARMINTERNALIDHASHTABLE : COL.IMap2;
	_HASHTABLEFACTORY : COL.HashTableFactory;
	_UDINTELEMFACTORY : COL.UdintElementFactory;
	_ULINTELEMFACTORY : COL.UlintElementFactory;
END_VAR
END_FUNCTION_BLOCK

METHOD FB_EXIT : BOOL
VAR_INPUT
	BINCOPYCODE : BOOL;
END_VAR
END_METHOD

METHOD FINDALARM : POINTER TO Alarm
VAR_INPUT
	UDIID : UDINT;
END_VAR
END_METHOD

METHOD FINDALARM2 : POINTER TO Alarm
VAR_INPUT
	UIID : ALARM_ID;
END_VAR
END_METHOD

METHOD FINDEVENT : POINTER TO Alarm
VAR_INPUT
	UIID : ALARM_ID;
END_VAR
END_METHOD

METHOD GETALARMSTORAGE : IDatabaseFileAlarmStorage
END_METHOD

METHOD GETTEXTLISTNAME2 : POINTER TO STRING
VAR_INPUT
	UIID : ALARM_ID;
END_VAR
END_METHOD

METHOD GETTEXTID : STRING
VAR_INPUT
	UIID : ALARM_ID;
	IWHICHMESSAGE : INT;
END_VAR
END_METHOD

METHOD GETID : ALARMGROUP_ID
END_METHOD

METHOD SETID
VAR_INPUT
	USIALARMGROUPID : ALARMGROUP_ID;
END_VAR
END_METHOD

METHOD GETSTRINGID2 : STRING
VAR_INPUT
	UDIALARMID : UDINT;
	IWHICHMESSAGE : INT;
END_VAR
VAR_OUTPUT
	STEXTID : STRING;
END_VAR
END_METHOD

METHOD RAISEEVENT2 : BOOL
VAR_INPUT
	EVENT : AlarmEvent;
END_VAR
VAR_OUTPUT
	ITFALARM : IAlarm;
END_VAR
END_METHOD

METHOD TRAVERSEALLALARMS
VAR_INPUT
	IWHICHALARMGROUP : INT;
	ITFALARMTRAVERSALCONSUMER : IAlarmTraversalConsumer;
END_VAR
END_METHOD

METHOD GETALARMS : POINTER TO ARRAY [0..0] OF Alarm
VAR_OUTPUT
	IALARMCOUNT : INT;
END_VAR
END_METHOD

METHOD GETEVENTS : POINTER TO ARRAY [0..0] OF Alarm
VAR_OUTPUT
	IEVENTCOUNT : INT;
END_VAR
END_METHOD

METHOD GETINTERNALID : UDINT
END_METHOD

METHOD GETNAME : STRING
END_METHOD

METHOD GETSTRINGID : STRING
VAR_INPUT
	UIID : ALARM_ID;
END_VAR
END_METHOD

METHOD GETTEXTLISTNAME : POINTER TO STRING
END_METHOD

METHOD GETVALUEPROVIDER : IValueProvider
END_METHOD

METHOD ISDEACTIVATED : BOOL
END_METHOD

METHOD RAISEEVENT : BOOL
VAR_INPUT
	EVENT : AlarmEvent;
END_VAR
END_METHOD

METHOD SETACTIVEALARM
VAR_INPUT
	IINDEX : INT;
	PALARM : POINTER TO Alarm;
END_VAR
END_METHOD

METHOD SETACTIVEALARMCOUNT
VAR_INPUT
	ICOUNT : INT;
END_VAR
END_METHOD

(* ---- ALARMGROUPADAPTER.fb ---- *)
FUNCTION_BLOCK ALARMGROUPADAPTER EXTENDS AlarmGroupContainerBase
END_FUNCTION_BLOCK

(* ---- ALARMGROUPCONTAINERBASE.fb ---- *)
FUNCTION_BLOCK ALARMGROUPCONTAINERBASE
VAR_INPUT
	M_SSTRINGID : STRING;
	M_STEXTLISTNAME : STRING;
	M_UDIINTERNALID : UDINT;
	M_SNAME : STRING;
END_VAR
END_FUNCTION_BLOCK

METHOD GETINTERNALID : UDINT
END_METHOD

METHOD GETNAME : STRING
END_METHOD

METHOD GETSTRINGID : STRING
VAR_INPUT
	UIID : ALARM_ID;
END_VAR
END_METHOD

METHOD GETTEXTLISTNAME : POINTER TO STRING
END_METHOD

METHOD FINDALARM : POINTER TO Alarm
VAR_INPUT
	UDIID : UDINT;
END_VAR
END_METHOD

METHOD FINDALARM2 : POINTER TO Alarm
VAR_INPUT
	UIID : ALARM_ID;
END_VAR
END_METHOD

METHOD GETALARMSTORAGE : IDatabaseFileAlarmStorage
END_METHOD

METHOD GETALARMS : POINTER TO ARRAY [0..0] OF Alarm
VAR_OUTPUT
	IALARMCOUNT : INT;
END_VAR
END_METHOD

METHOD GETEVENTS : POINTER TO ARRAY [0..0] OF Alarm
VAR_OUTPUT
	IEVENTCOUNT : INT;
END_VAR
END_METHOD

METHOD GETVALUEPROVIDER : IValueProvider
END_METHOD

METHOD ISDEACTIVATED : BOOL
END_METHOD

METHOD RAISEEVENT : BOOL
VAR_INPUT
	EVENT : AlarmEvent;
END_VAR
END_METHOD

METHOD SETACTIVEALARM
VAR_INPUT
	IINDEX : INT;
	PALARM : POINTER TO Alarm;
END_VAR
END_METHOD

METHOD SETACTIVEALARMCOUNT
VAR_INPUT
	ICOUNT : INT;
END_VAR
END_METHOD

(* ---- ALARMGROUPMOCK.fb ---- *)
FUNCTION_BLOCK ALARMGROUPMOCK EXTENDS AlarmGroupContainerBase
END_FUNCTION_BLOCK

METHOD SETVALUES
VAR_INPUT
	ISET : INT;
END_VAR
END_METHOD

(* ---- ALARMINSTANCEDICTIONARY.fb ---- *)
FUNCTION_BLOCK ALARMINSTANCEDICTIONARY
VAR
	_ALARMINSTANCEHASHTABLE : COL.IMap2 := NULL;
	_HASHTABLEFACTORY : COL.HashTableFactory;
	_HASHTABLEVALUEELEMFACTORY : HashtableValueElementFactory;
	_HASHTABLEKEYELEMFACTORY : HashtableKeyElementFactory;
END_VAR
END_FUNCTION_BLOCK

METHOD ADDINSTANCE : COL.COLLECTION_ERROR
VAR_INPUT
	PINSTANCE : POINTER TO BYTE;
	PSTALARMTEMPLATENAME : POINTER TO STRING;
	UDIALARMGROUPID : UDINT;
	UITEMPLATEALARMSOFFSET : UINT;
	UITEMPLATEALARMSLENGTH : UINT;
	UITEMPLATEEVENTSOFFSET : UINT;
	UITEMPLATEEVENTSLENGTH : UINT;
END_VAR
END_METHOD

METHOD CLEARALLOFALARMGROUP : BOOL
END_METHOD

METHOD GETINSTANCE : IHashtableValueElement
VAR_INPUT
	PINSTANCE : POINTER TO BYTE;
	UDIALARMID : REFERENCE TO ALARM_ID;
	STALARMTEMPLATENAME : REFERENCE TO STRING;
END_VAR
END_METHOD

METHOD PRVCREATEKEYELEMENT : IHashtableKeyElement
VAR_INPUT
	PINSTANCE : POINTER TO BYTE;
	PSTALARMTEMPLATENAME : POINTER TO STRING;
END_VAR
VAR_OUTPUT
	FBFERROR : COL.FBF.ERROR;
END_VAR
END_METHOD

(* ---- ALARMLATCHADAPTER.fb ---- *)
FUNCTION_BLOCK ALARMLATCHADAPTER
VAR
	_ALARMLATCH : IAlarmMetaObjectStubSupportsAdditionalLatchVariables;
END_VAR
END_FUNCTION_BLOCK

METHOD FB_INIT : BOOL
VAR_INPUT
	BINITRETAINS : BOOL;
	BINCOPYCODE : BOOL;
	ALARMLATCH : IAlarmMetaObjectStub3;
END_VAR
END_METHOD

METHOD GETCOUNTLATCHVARIABLES : USINT
END_METHOD

METHOD GETLATCHVARVALUE : AlarmManager_Interfaces.ITypedValue
VAR_INPUT
	IWHICHLATCHVAR : INT;
END_VAR
END_METHOD

METHOD INITIALIZE : BOOL
VAR_INPUT
	ALARMLATCH : IAlarmMetaObjectStubSupportsAdditionalLatchVariables;
END_VAR
END_METHOD

METHOD SETLATCHVARVALUE
VAR_INPUT
	IWHICHLATCHVAR : INT;
	ITFTYPEDVALUELATCHVAR : AlarmManager_Interfaces.ITypedValue;
END_VAR
END_METHOD

(* ---- ALARMMANAGERCLIENTINFOSTRUCTVECTOR.fb ---- *)
FUNCTION_BLOCK ALARMMANAGERCLIENTINFOSTRUCTVECTOR EXTENDS BaseVector
VAR
	_PARRALARMMANAGERCLIENTINFOSTRUCT : POINTER TO ARRAY [0..MAX_NUM_ENTRIES] OF POINTER TO AlarmManagerClientInfoStruct;
	MAX_NUM_ENTRIES : INT := 10;
END_VAR
END_FUNCTION_BLOCK

METHOD ABSTRASSIGN : UDINT
VAR_INPUT
	PBT : POINTER TO BYTE;
	UDIINDEX : UDINT;
END_VAR
END_METHOD

METHOD ABSTRDATAPTRCHANGED : UDINT
END_METHOD

METHOD ABSTRSIZEOFELEMENT : UDINT
END_METHOD

METHOD PRVFINDALARMMANAGERCLIENTINFOSTRUCT : UDINT
VAR_INPUT
	ITFALARMMANAGERCLIENT : IAlarmManagerClient;
END_VAR
VAR_OUTPUT
	UDIRESULT : UDINT;
END_VAR
END_METHOD

METHOD ADDALARMMANAGERCLIENTINFOSTRUCT : UDINT
VAR_INPUT
	PITEM : POINTER TO AlarmManagerClientInfoStruct;
END_VAR
END_METHOD

METHOD GETALARMMANAGERCLIENTINFOSTRUCT : POINTER TO AlarmManagerClientInfoStruct
VAR_INPUT
	ITFALARMMANAGERCLIENT : IAlarmManagerClient;
END_VAR
VAR_OUTPUT
	UDIRESULT : UDINT;
END_VAR
END_METHOD

METHOD GETALARMMANAGERCLIENTINFOSTRUCTAT : POINTER TO AlarmManagerClientInfoStruct
VAR_INPUT
	UDIINDEX : UDINT;
END_VAR
VAR_OUTPUT
	UDIRESULT : UDINT;
END_VAR
END_METHOD

METHOD REMOVEALARMMANAGERCLIENTINFOSTRUCT : UDINT
VAR_INPUT
	ITFALARMMANAGERCLIENT : IAlarmManagerClient;
END_VAR
END_METHOD

(* ---- ALARMMANAGERREALVALUESTATISTICS.fb ---- *)
FUNCTION_BLOCK ALARMMANAGERREALVALUESTATISTICS
VAR_OUTPUT
	RAVG : REAL;
	RSTDDERIV : REAL;
	RMIN : REAL := 3.402823466E+38;
	RMAX : REAL := -3.402823466E+38;
	UDINUM : UDINT;
END_VAR
VAR
	RM2 : REAL;
END_VAR
END_FUNCTION_BLOCK

METHOD ADDVALUE
VAR_INPUT
	RVALUE : REAL;
END_VAR
END_METHOD

METHOD RESET
END_METHOD

(* ---- ALARMMOCK.fb ---- *)
FUNCTION_BLOCK ALARMMOCK EXTENDS AlarmContainerBase
VAR
	M_ALARMGROUP : AlarmGroupMock;
	M_ALARMCLASS : AlarmClassMock;
END_VAR
END_FUNCTION_BLOCK

METHOD FB_EXIT : BOOL
VAR_INPUT
	BINCOPYCODE : BOOL;
END_VAR
END_METHOD

METHOD FB_INIT : BOOL
VAR_INPUT
	BINITRETAINS : BOOL;
	BINCOPYCODE : BOOL;
END_VAR
END_METHOD

METHOD SETVALUES
VAR_INPUT
	ISET : INT;
END_VAR
END_METHOD

METHOD GETCURRENTVALUE : AlarmManager_Interfaces.ITypedValue
END_METHOD

METHOD GETLATCHVARVALUE : ITypedValue
VAR_INPUT
	IWHICHLATCHVAR : INT;
END_VAR
END_METHOD

METHOD GETTRIGGERVALUE : AlarmManager_Interfaces.ITypedValue
END_METHOD

(* ---- ALARMROOTPAGEREADWRITEMODEPROVIDER.fb ---- *)
FUNCTION_BLOCK ALARMROOTPAGEREADWRITEMODEPROVIDER
VAR
	M_XREADONLY : BOOL;
	M_HSEM : RTS_IEC_HANDLE := RTS_INVALID_HANDLE;
	READONLY : BOOL;
END_VAR
END_FUNCTION_BLOCK

METHOD FB_EXIT : BOOL
VAR_INPUT
	BINCOPYCODE : BOOL;
END_VAR
END_METHOD

METHOD FB_INIT : BOOL
VAR_INPUT
	BINITRETAINS : BOOL;
	BINCOPYCODE : BOOL;
END_VAR
END_METHOD

(* ---- ALARMSERVICEALARMSTORAGEREADERCONSUMER.fb ---- *)
FUNCTION_BLOCK ALARMSERVICEALARMSTORAGEREADERCONSUMER
VAR
	M_IMAXCOUNTROWSTOREAD : INT;
	M_USICOUNTLATCHVARIABLES : USINT;
	M_IEFFECTIVENUMBEROFROWS : INT;
	M_PAALARMSTORAGESTATICDATA : POINTER TO ARRAY [0..0] OF AlarmStorageStaticData;
	M_PALATCHVARIABLES : POINTER TO ARRAY [0..0] OF AlarmStorageLatchVariable;
	M_IEFFECTIVEARRAYSIZE : INT;
	COMPONENT : STRING := 'AlarmServiceAlarmStorageReaderConsumer';
END_VAR
END_FUNCTION_BLOCK

METHOD FB_EXIT : BOOL
VAR_INPUT
	BINCOPYCODE : BOOL;
END_VAR
END_METHOD

METHOD GETALARM : AlarmStorageStaticData
VAR_INPUT
	IWHICHROW : INT;
END_VAR
END_METHOD

METHOD GETCOUNTLATCHVARIABLES : USINT
END_METHOD

METHOD GETCOUNTROWS : INT
END_METHOD

METHOD GETLATCHVARIABLE : AlarmStorageLatchVariable
VAR_INPUT
	IWHICHROW : INT;
	USIWHICHVARIABLE : USINT;
END_VAR
END_METHOD

METHOD INITIALIZE
VAR_INPUT
	IMAXCOUNTROWSTOREAD : INT;
END_VAR
END_METHOD

METHOD ALARMREAD
VAR_INPUT
	DIWHICHROW : DINT;
	STATICDATA : AlarmStorageStaticData;
END_VAR
END_METHOD

METHOD BEFOREREADING
VAR_INPUT
	USICOUNTLATCHVARIABLES : USINT;
END_VAR
END_METHOD

METHOD LATCHVARIABLEREAD
VAR_INPUT
	DIWHICHROW : DINT;
	USIWHICHVARIABLE : USINT;
	LILATCHVARVALUE : LINT;
	ILATCHVARTYPE : TypeClass;
	XVALUENULL : BOOL;
END_VAR
END_METHOD

METHOD READINGDATACOMPLETED
END_METHOD

METHOD PRVFREEBUFFERS
VAR_INPUT
	XFREESTATICDATA : BOOL;
	XFREELATCHVARIABLES : BOOL;
END_VAR
END_METHOD

(* ---- ALARMSERVICEHANDLER.fb ---- *)
FUNCTION_BLOCK ALARMSERVICEHANDLER
VAR
	_HBTR : RTS_IEC_HANDLE := RTS_INVALID_HANDLE;
	_HBTW : RTS_IEC_HANDLE := RTS_INVALID_HANDLE;
	_PCURRENTCONTENT : POINTER TO BYTE;
	_UDICURRENTCONTENTLENGTH : UDINT;
	_UDIPOSITION : UDINT;
	_CURRENTTAGTYPE : CmpBinTagUtilIec.BTagElementType;
	_TARGETBYTEORDER : EAlarmByteOrder := AlarmFctGetLocalByteorder();
	_UDIBUFFERSIZE : UDINT;
	_FILTERCRITERIA : VisuFbAlarmFilterCriteriaService;
	_ALARMSERVICEHANDLERBUFFERPROVIDER : AlarmServiceHandlerBufferProvider;
	_RESULTDATABLOCK : BinTagWriterDataBlock;
	_UDIRESULT : UDINT;
	_UISERVICE : UINT;
	_ITFALARMTRAVERSALCONSUMER : IAlarmTraversalConsumer := THIS^;
	_ARRALARMGROUPRECORD : ARRAY [0..(MAX_GROUP_RECORD - 1)] OF AlarmRecord;
	_IRECORDIDPROGRESSIVE : INT;
	_PBYTESBUFFER : POINTER TO BYTE;
	_ALARMMOCK : AlarmMock;
	_ALARMGROUPMOCK : AlarmGroupMock;
	_ALARMCLASSMOCK : AlarmClassMock;
	_HISTORICALALARMMOCK : HistoricalAlarmMock;
	_DIACTIVEALMCNT : DINT;
	_IRECORDID : INT;
	_AROWID : ARRAY [1..SIZE_HIST_ACTIVE_ALM] OF HistoricalActiveAlarmRowID;
	_IROWIDPROGCOUNT : INT;
	_XBUFFEROVERMSG : BOOL;
	_LASTSTORAGECLEARVALUE : INT := INITIAL_VALUE;
	_LASTSTORAGECOUNTER : DINT := INITIAL_VALUE;
	_CACHEDHISTORICROWCOUNT : DINT;
	BYTE_BUFFER_SIZE : INT := 4096;
	COMPONENT : STRING := 'AlarmServiceHandler';
	MAX_GROUP_RECORD : INT := 25;
	INITIAL_VALUE : INT := 0;
END_VAR
END_FUNCTION_BLOCK

METHOD FB_EXIT : BOOL
VAR_INPUT
	BINCOPYCODE : BOOL;
END_VAR
END_METHOD

METHOD FB_INIT : BOOL
VAR_INPUT
	BINITRETAINS : BOOL;
	BINCOPYCODE : BOOL;
END_VAR
END_METHOD

METHOD HANDLEEVENTS : UDINT
VAR_INPUT
	IEVENT : INT;
	PEVENTPARAM : POINTER TO BYTE;
END_VAR
END_METHOD

METHOD HANDLESERVICE : UDINT
VAR_INPUT
	PPARAMETERS : POINTER TO SERVICEHANDLER_PARAMETER;
END_VAR
END_METHOD

METHOD AFTERLASTALARMOFALARMGROUP
VAR_INPUT
	ITFALARMGROUP : IAlarmGroup;
END_VAR
END_METHOD

METHOD ALARMCLASSREACHED
VAR_INPUT
	ITFALARMCLASS : IAlarmClass;
END_VAR
END_METHOD

METHOD ALARMHISTORICALISRELEVANT : BOOL
VAR_INPUT
	ROW : REFERENCE TO AlarmStorageRow;
END_VAR
END_METHOD

METHOD ALARMHISTORICALREACHED : UDINT
VAR_INPUT
	ROW : REFERENCE TO AlarmStorageRow;
END_VAR
END_METHOD

METHOD ALARMREACHED
VAR_INPUT
	IWHICHALARMGROUP : INT;
	IWHICHALARM : INT;
	ITFALARM : IAlarm3;
END_VAR
END_METHOD

METHOD BEFOREFIRSTALARMOFALARMGROUP
VAR_INPUT
	ITFALARMGROUP : IAlarmGroup;
END_VAR
END_METHOD

METHOD BEGINTRAVERSAL
END_METHOD

METHOD ENDTRAVERSAL
END_METHOD

METHOD GETACTIVEALARMHISTORICALROWID
VAR_INPUT
	XFIRST : BOOL;
END_VAR
VAR_OUTPUT
	DWROWID : DWORD;
	LITS : LINT;
END_VAR
END_METHOD

METHOD WRITEBYTE : UDINT
VAR_INPUT
	BT : BYTE;
END_VAR
END_METHOD

METHOD WRITECOMPLEXSTARTTAG : UDINT
VAR_INPUT
	UDITAG : UDINT;
	UDIMINLENSIZE : UDINT;
END_VAR
END_METHOD

METHOD WRITEDWORD : UDINT
VAR_INPUT
	DW : DWORD;
END_VAR
END_METHOD

METHOD WRITEDATASTARTTAG : UDINT
VAR_INPUT
	UDITAG : UDINT;
	ALIGNMENT : CmpBinTagUtilIec.BTagAlignment;
	UDIMINLENSIZE : UDINT;
END_VAR
END_METHOD

METHOD WRITEENDTAG : UDINT
VAR_INPUT
	UDITAG : UDINT;
END_VAR
END_METHOD

METHOD WRITEFILLBYTES : UDINT
END_METHOD

METHOD WRITELWORD : UDINT
VAR_INPUT
	LW : LWORD;
END_VAR
END_METHOD

METHOD WRITESTRING : UDINT
VAR_INPUT
	PSSTRING : POINTER TO STRING(255);
END_VAR
END_METHOD

METHOD WRITEWSTRING : UDINT
VAR_INPUT
	PWSSTRING : POINTER TO WSTRING(255);
END_VAR
END_METHOD

METHOD WRITEWORD : UDINT
VAR_INPUT
	WD : WORD;
END_VAR
END_METHOD

METHOD PRVACKNOWLEDGE : UDINT
VAR_INPUT
	PPARAMETERS : POINTER TO SERVICEHANDLER_PARAMETER;
END_VAR
END_METHOD

METHOD PRVCHANNELTEST : UDINT
VAR_INPUT
	PPARAMETERS : POINTER TO SERVICEHANDLER_PARAMETER;
END_VAR
END_METHOD

METHOD PRVGETALARMS : UDINT
VAR_INPUT
	PPARAMETERS : POINTER TO SERVICEHANDLER_PARAMETER;
END_VAR
END_METHOD

METHOD PRVGETALARMS2 : UDINT
VAR_INPUT
	PPARAMETERS : POINTER TO SERVICEHANDLER_PARAMETER;
END_VAR
END_METHOD

METHOD PRVGETALARMS3 : UDINT
VAR_INPUT
	PPARAMETERS : POINTER TO SERVICEHANDLER_PARAMETER;
END_VAR
END_METHOD

METHOD PRVGETCOUNTALARMS : UDINT
VAR_INPUT
	PPARAMETERS : POINTER TO SERVICEHANDLER_PARAMETER;
END_VAR
END_METHOD

METHOD PRVGETMINMAXTIMESTAMPS : UDINT
VAR_INPUT
	PPARAMETERS : POINTER TO SERVICEHANDLER_PARAMETER;
END_VAR
END_METHOD

METHOD PRVGETTYPEDVALUE
VAR_INPUT
	ITFTYPEDVALUE : ITypedValue;
END_VAR
VAR_OUTPUT
	BYTYPECLASS : BYTE;
	LIVALUE : LINT;
END_VAR
END_METHOD

METHOD PRVGETACTIVEALARMS : UDINT
VAR_INPUT
	PPARAMETERS : POINTER TO SERVICEHANDLER_PARAMETER;
END_VAR
END_METHOD

METHOD PRVGETACTIVEALARMS2 : UDINT
VAR_INPUT
	PPARAMETERS : POINTER TO SERVICEHANDLER_PARAMETER;
END_VAR
END_METHOD

METHOD PRVGETACTIVEALARMSALARMREACHED
VAR_INPUT
	ITFALARM : IAlarm3;
	UISERVICE : UINT;
END_VAR
END_METHOD

METHOD PRVGETALARMCLASSCONFIGURATION : UDINT
VAR_INPUT
	PPARAMETERS : POINTER TO SERVICEHANDLER_PARAMETER;
END_VAR
END_METHOD

METHOD PRVGETALARMCONFIGURATION : UDINT
VAR_INPUT
	PPARAMETERS : POINTER TO SERVICEHANDLER_PARAMETER;
END_VAR
END_METHOD

METHOD PRVGETALARMCONFIGURATION2 : UDINT
VAR_INPUT
	PPARAMETERS : POINTER TO SERVICEHANDLER_PARAMETER;
END_VAR
END_METHOD

METHOD PRVGETALARMCONFIGURATIONAFTERLASTALARMOFALARMGROUP
VAR_INPUT
	ITFALARMGROUP : IAlarmGroup;
END_VAR
END_METHOD

METHOD PRVGETALARMCONFIGURATIONALARMCLASSREACHED
VAR_INPUT
	ITFALARMCLASS : IAlarmClass;
END_VAR
END_METHOD

METHOD PRVGETALARMCONFIGURATIONALARMREACHED
VAR_INPUT
	IWHICHALARMGROUP : INT;
	IWHICHALARM : INT;
	ITFALARM : IAlarm3;
	UISERVICE : UINT;
END_VAR
END_METHOD

METHOD PRVGETALARMCONFIGURATIONBEFOREFIRSTALARMOFALARMGROUP
VAR_INPUT
	ITFALARMGROUP : IAlarmGroup;
END_VAR
END_METHOD

METHOD PRVRESETALARMSRECORD : UDINT
VAR_INPUT
	PPARAMETERS : POINTER TO SERVICEHANDLER_PARAMETER;
END_VAR
END_METHOD

METHOD PRVSETALARMSRECORD : UDINT
VAR_INPUT
	PPARAMETERS : POINTER TO SERVICEHANDLER_PARAMETER;
END_VAR
END_METHOD

METHOD PRVSETALARMSRECORDALARMCLASSREACHED
VAR_INPUT
	ITFALARMCLASS : IAlarmClass;
END_VAR
END_METHOD

METHOD PRVFILLFILTERCRITERIA : BOOL
VAR_INPUT
	UDITAGID : UDINT;
END_VAR
VAR_OUTPUT
	UDIRESULT : UDINT;
END_VAR
END_METHOD

METHOD PRVFILLLATCHFILTERCRITERIA : UDINT
END_METHOD

METHOD PRVFILLTIMERANGEFILTERCRITERIA : UDINT
END_METHOD

METHOD PRVINITIALIZEFILTERCRITERIA
END_METHOD

METHOD PRVGETACTIVEALARMHISTORICALROWID
VAR_INPUT
	XFIRST : BOOL;
END_VAR
VAR_OUTPUT
	DWROWID : DWORD;
	LITS : LINT;
END_VAR
END_METHOD

METHOD PRVGETHISTORICALACTIVEALARMS : UDINT
VAR_INPUT
	PPARAMETERS : POINTER TO SERVICEHANDLER_PARAMETER;
END_VAR
END_METHOD

METHOD PRVGETHISTORICALACTIVEALARMSREACHED : UDINT
VAR_INPUT
	ROW : REFERENCE TO AlarmStorageRow;
END_VAR
END_METHOD

METHOD PRVGETHISTORICALALARMS : UDINT
VAR_INPUT
	PPARAMETERS : POINTER TO SERVICEHANDLER_PARAMETER;
END_VAR
END_METHOD

METHOD PRVGETHISTORICALALARMSCONFIG : UDINT
VAR_INPUT
	PPARAMETERS : POINTER TO SERVICEHANDLER_PARAMETER;
END_VAR
END_METHOD

METHOD PRVGETHISTORICALALARMSISRELEVANT : BOOL
VAR_INPUT
	ROW : REFERENCE TO AlarmStorageRow;
END_VAR
END_METHOD

METHOD PRVGETHISTORICALALARMSREACHED : UDINT
VAR_INPUT
	ROW : REFERENCE TO AlarmStorageRow;
END_VAR
END_METHOD

METHOD PRVGETROWCOUNT : DINT
END_METHOD

METHOD PRVCREATEDYNAMIC : UDINT
VAR_INPUT
	PDATABUFFERREADER : POINTER TO BYTE;
	UDIDATABUFFERREADERSIZE : UDINT;
	PDATABUFFERWRITER : POINTER TO BYTE;
	UDIDATABUFFERWRITERSIZE : UDINT;
END_VAR
END_METHOD

METHOD PRVDESTROY : UDINT
END_METHOD

METHOD PRVINIT : UDINT
VAR_INPUT
	PDATABUFFERREADER : POINTER TO BYTE;
	UDIDATABUFFERREADERSIZE : UDINT;
	PDATABUFFERWRITER : POINTER TO BYTE;
	UDIDATABUFFERWRITERSIZE : UDINT;
END_VAR
END_METHOD

METHOD PRVISDATATAG : BOOL
END_METHOD

METHOD PRVISOURAPPLICATION : BOOL
VAR_INPUT
	SAPPLICATIONNAME : STRING;
END_VAR
END_METHOD

METHOD PRVISTOPLEVEL : BOOL
END_METHOD

METHOD PRVMOVEDOWN : UDINT
END_METHOD

METHOD PRVMOVENEXT : UDINT
END_METHOD

METHOD PRVMOVENEXTCONDITIONAL : UDINT
VAR_INPUT
	XDOMOVE : BOOL;
END_VAR
END_METHOD

METHOD PRVMOVEUP : UDINT
END_METHOD

METHOD PRVREADBYTE : UDINT
VAR_OUTPUT
	BT : BYTE;
END_VAR
END_METHOD

METHOD PRVREADBYTES : UDINT
VAR_INPUT
	UDISIZE : UDINT;
	PBYTE : POINTER TO BYTE;
END_VAR
END_METHOD

METHOD PRVREADDWORD : UDINT
VAR_OUTPUT
	DW : DWORD;
END_VAR
END_METHOD

METHOD PRVREADLWORD : UDINT
VAR_OUTPUT
	LW : LWORD;
END_VAR
END_METHOD

METHOD PRVREADSTARTTAG : UDINT
END_METHOD

METHOD PRVREADSTRING : UDINT
VAR_OUTPUT
	STR : STRING(255);
END_VAR
END_METHOD

METHOD PRVREADWORD : UDINT
VAR_OUTPUT
	WD : WORD;
END_VAR
END_METHOD

METHOD PRVWRITEBYTES : UDINT
VAR_INPUT
	PDATA : POINTER TO BYTE;
	UDISIZE : UDINT;
END_VAR
END_METHOD

METHOD PRVWRITESTRING : UDINT
VAR_INPUT
	STR : STRING(255);
END_VAR
END_METHOD

METHOD PRVALMRECORDADDALARMCLASSES : BOOL
VAR_INPUT
	IRECORDID : INT;
	ITFALARMCLASS : IAlarmClass;
END_VAR
END_METHOD

METHOD PRVALMRECORDADDNEWALARMCLASSES : BOOL
VAR_INPUT
	IRECORDID : INT;
	ICLASS : INT;
END_VAR
END_METHOD

METHOD PRVALMRECORDCREATERECORD : POINTER TO AlarmRecord
VAR_INPUT
	IGROUP : INT;
END_VAR
END_METHOD

METHOD PRVALMRECORDDISPLAYSTATUS
END_METHOD

METHOD PRVALMRECORDFREEAREAS
VAR_INPUT
	IX : INT;
END_VAR
END_METHOD

METHOD PRVALMRECORDGETRECORD : POINTER TO AlarmRecord
VAR_INPUT
	IRECORDID : INT;
END_VAR
END_METHOD

METHOD PRVALMRECORDREMOVE : INT
VAR_INPUT
	IRECORDID : INT;
END_VAR
END_METHOD

METHOD PRVALMRECORDREMOVEALL
END_METHOD

METHOD PRVALMRECORDREMOVECLIENT : INT
VAR_INPUT
	UICLIENT : UINT;
END_VAR
END_METHOD

(* ---- ALARMSERVICEHANDLERBUFFERPROVIDER.fb ---- *)
FUNCTION_BLOCK ALARMSERVICEHANDLERBUFFERPROVIDER
VAR
	M_PAUDIALARMGROUPS : POINTER TO ARRAY [0..0] OF UDINT;
	M_PAUDIALARMCLASSES : POINTER TO ARRAY [0..0] OF UDINT;
	M_PALATCHVARIABLES : POINTER TO ARRAY [0..0] OF LatchVariable;
	M_PAALARMSTOACKBUFFER : POINTER TO ARRAY [0..0] OF AlarmToAcknowledge;
	M_ICOUNTALARMGROUPS : INT;
	M_ICOUNTALARMCLASSES : INT;
	M_ICOUNTLATCHVARIABLES : INT;
	M_ICOUNTALARMSTOACK : INT;
	COMPONENT : STRING := 'AlarmFilterCriteriaBufferProvider';
END_VAR
END_FUNCTION_BLOCK

METHOD ALLOCATEALARMCLASSFILTERBUFFER : POINTER TO ARRAY [0..0] OF UDINT
VAR_INPUT
	IREQUIREDMINIMUMSIZE : INT;
END_VAR
END_METHOD

METHOD ALLOCATEALARMGROUPFILTERBUFFER : POINTER TO ARRAY [0..0] OF UDINT
VAR_INPUT
	IREQUIREDMINIMUMSIZE : INT;
END_VAR
END_METHOD

METHOD ALLOCATEALARMSTOACKBUFFER : POINTER TO ARRAY [0..0] OF AlarmToAcknowledge
VAR_INPUT
	IREQUIREDMINIMUMSIZE : INT;
END_VAR
END_METHOD

METHOD ALLOCATELATCHVARIABLESBUFFER : POINTER TO ARRAY [0..0] OF LatchVariable
VAR_INPUT
	IREQUIREDMINIMUMSIZE : INT;
END_VAR
END_METHOD

METHOD FB_EXIT : BOOL
VAR_INPUT
	BINCOPYCODE : BOOL;
END_VAR
END_METHOD

METHOD FREEBUFFERS
VAR_INPUT
	XFREEALARMGROUPSBUFFER : BOOL;
	XFREEALARMCLASSESBUFFER : BOOL;
	XFREELATCHVARIABLES : BOOL;
	XFREEALARMSTOACKBUFFER : BOOL;
END_VAR
END_METHOD

(* ---- ALARMSTATECHANGEDEVENTLISTENER.fb ---- *)
FUNCTION_BLOCK ALARMSTATECHANGEDEVENTLISTENER
VAR
	_ITFALARMSTATECHANGEDLISTENERS : ARRAY [0..4] OF IAlarmStateChangedListener := [NULL, NULL, NULL, NULL, NULL];
END_VAR
END_FUNCTION_BLOCK

METHOD ACTIONSTATECHANGED : BOOL
VAR_INPUT
	ITFALARM : IAlarm;
	ESTATEOLD : AlarmState;
	ESTATENEW : AlarmState;
	ESTATETRANSITION : AlarmStateTransition;
END_VAR
END_METHOD

METHOD DEACTIVATIONSTATECHANGED : BOOL
VAR_INPUT
	ITFALARM : IAlarm;
	XNEWDEACTIVATIONSTATE : BOOL;
END_VAR
END_METHOD

METHOD REGISTERLISTENER : BOOL
VAR_INPUT
	ITFALARMSTATECHANGEDLISTENER : IAlarmStateChangedListener;
END_VAR
END_METHOD

(* ---- ALARMSTORAGELIMIT.fb ---- *)
FUNCTION_BLOCK ALARMSTORAGELIMIT
VAR_INPUT
	_UXILIMIT : CAA.COUNT;
END_VAR
VAR
	_UXICURRENT : CAA.COUNT;
	_LIMITASSIGNED : BOOL;
	ACTIVE : BOOL;
END_VAR
END_FUNCTION_BLOCK

METHOD CANINCREMENT : BOOL
VAR_INPUT
	UXIADDITIONALALARMS : CAA.COUNT;
END_VAR
END_METHOD

METHOD DECREMENT
VAR_INPUT
	COUNT : CAA.COUNT;
END_VAR
END_METHOD

METHOD INCREMENT
VAR_INPUT
	COUNT : CAA.COUNT;
END_VAR
END_METHOD

METHOD SETLIMIT : BOOL
VAR_INPUT
	UXILIMIT : CAA.COUNT;
END_VAR
END_METHOD

(* ---- ALARMSTORAGELOCALBUFFERACCESS.fb ---- *)
FUNCTION_BLOCK ALARMSTORAGELOCALBUFFERACCESS EXTENDS AbstractDatabaseAccess
VAR
	M_CONTEXT : LocalBufferDatabaseAccessContext;
	M_ECURRSTATE : EAlarmStorageMirrorState;
	M_XCURRENTMIRRORINGINVALID : BOOL;
	M_ALARMSTORAGEREADER : AlarmStorageReader;
	M_LIMINTIMESTAMP : LINT;
	M_LIMAXTIMESTAMP : LINT;
	M_UDICOUNTALARMS : UDINT;
	M_UDICOUNTLATCHVARIABLES : UDINT;
	M_PALIBUFFER : POINTER TO ARRAY [0..0] OF LINT;
	M_UDIBUFFERSIZE : UDINT;
	M_UDIMAXROWCOUNT : UDINT;
	M_UXIROWCOUNT : CAA.COUNT;
	M_PADIINDEXMAPPINGBUFFER : POINTER TO ARRAY [0..100] OF DINT;
	M_UDIINDEXMAPPINGBUFFERSIZE : UDINT;
	M_DICIRCULARBUFFERBORDER : DINT;
	M_XCIRCULARBUFFER : BOOL;
	M_UDICOUNTBYTESPERALARM : UDINT;
	M_DIALARMINDEX : DINT;
	M_PALICURRALARM : POINTER TO ARRAY [0..0] OF LINT;
	M_UDIOFFSETTRIGGERVALUETYPE : UDINT;
	M_XADDEDASALARMSTORAGELISTENER : BOOL;
	M_TSLASTCOMPARER : TSLastComparer;
	M_TSACTIVECOMPARER : TSActiveComparer;
	M_TSINACTIVECOMPARER : TSInactiveComparer;
	M_TSACKCOMPARER : TSAckComparer;
	M_PRIORITYCOMPARER : PriorityComparer;
	M_STATECOMPARER : StateComparer;
	M_ALARMCLASSCOMPARER : AlarmClassComparer;
	M_MESSAGECOMPARER : MessageComparer;
	M_VALUECOMPARER : ValueComparer;
	M_REMOTEDEVICECOMPARER : RemoteDeviceComparer;
	M_COMMENTACKCOMPARER : CommentComparer;
	M_USERIDACKCOMPARER : UserIdComparer;
	M_AITFALARMSTORAGEDATACOMPARER : ARRAY [EAlarmComparable.FIRST_ENTRY..EAlarmComparable.LAST_ENTRY] OF IAlarmStorageDataComparer;
	M_ITFALARMSTORAGEDATACOMPARER : IAlarmStorageDataComparer := m_TSLastComparer;
	M_XSORTASCENDING : BOOL := FALSE;
	M_XSORTREQUIRED : BOOL;
	M_ITFMEMORYMANAGER : AlarmManagerInternal_Interfaces.IMemoryManager;
	M_ITFALARMSTORAGEREADERCONSUMER : IAlarmStorageReaderConsumer := THIS^;
	M_ITFALARMSTORAGELISTENER : IAlarmStorageListener := THIS^;
	M_ITFRANDOMALARMREADACCESS : IRandomAlarmReadAccess := THIS^;
	M_HSEMSORTING : SysSem.RTS_IEC_HANDLE := SysSem.RTS_INVALID_HANDLE;
	M_XALARMCOUNTLIMITEXCEEDED : BOOL;
	COMPONENT : STRING := 'AlarmStorageLocalBufferAccess';
	M_STARTMIRRORING : LTIME;
	M_XDISPLAYDONE : BOOL;
	OFFSET_ROWID : UDINT := 0;
	OFFSET_GROUPID : UDINT := 4;
	OFFSET_CLASSID : UDINT := 8;
	OFFSET_ALARMID : UDINT := 12;
	OFFSET_TSLAST : UDINT := 16;
	OFFSET_TSACTIVE : UDINT := 24;
	OFFSET_TSINACTIVE : UDINT := 32;
	OFFSET_TSACK : UDINT := 40;
	OFFSET_OFFSETLAST : UDINT := 48;
	OFFSET_OFFSETACTIVE : UDINT := 50;
	OFFSET_OFFSETINACTIVE : UDINT := 52;
	OFFSET_OFFSETACKN : UDINT := 54;
	OFFSET_TVALUE : UDINT := 56;
	OFFSET_PRIORITY : UDINT := 64;
	OFFSET_STATE : UDINT := 65;
	OFFSET_REMOTEDEVICE : UDINT := 68;
	OFFSET_CMTACTIVEACK : UDINT := 80;
	OFFSET_USERIDACTIVEACK : UDINT := 88;
	OFFSET_CMTNORMAL : UDINT := 96;
	OFFSET_USERIDNORMAL : UDINT := 104;
	OFFSET_CMTACTIVE : UDINT := 112;
	OFFSET_USERIDACTIVE : UDINT := 120;
	OFFSET_CMTWAITINGCONF : UDINT := 128;
	OFFSET_USERIDWAITINGCONF : UDINT := 136;
	OFFSET_START_LATCHVARIABLES : UDINT := 144;
	SIZEOFVALUE : UDINT := 8;
	SIZEOFTYPE : UDINT := 1;
	SUPPORTED_VERSION : INT := DBVersions.LATEST_VERSION;
	ALARMCOUNTLIMITEXCEEDED : BOOL;
	BYTEORDER : EAlarmByteOrder;
END_VAR
END_FUNCTION_BLOCK

METHOD BEFOREPROCESSING
END_METHOD

METHOD CYCLICCALL : EAlarmStorageMirrorState
END_METHOD

METHOD FB_EXIT : BOOL
VAR_INPUT
	BINCOPYCODE : BOOL;
END_VAR
END_METHOD

METHOD FB_INIT : BOOL
VAR_INPUT
	BINITRETAINS : BOOL;
	BINCOPYCODE : BOOL;
END_VAR
END_METHOD

METHOD FILL : UDINT
END_METHOD

METHOD ISBUSY : BOOL
END_METHOD

METHOD REVERSEORDER
END_METHOD

METHOD SETMEMORYMANAGER
VAR_INPUT
	ITFMEMORYMANAGER : AlarmManagerInternal_Interfaces.IMemoryManager;
END_VAR
END_METHOD

METHOD SORTALARMS
VAR_INPUT
	EORDERCRITERION : EAlarmComparable;
	IWHICHCHARACTERISTIC : INT;
	STRINGTYPE : __SYSTEM.TYPE_CLASS;
	XSORTASCENDING : BOOL;
END_VAR
END_METHOD

METHOD ALARMADDED
VAR_INPUT
	ALARM : AlarmStorageRow;
END_VAR
END_METHOD

METHOD ALARMMODIFIED
VAR_INPUT
	ALARM : AlarmStorageRow;
END_VAR
END_METHOD

METHOD ALARMDELETED
VAR_INPUT
	IDROW : CAA.IDENT;
END_VAR
END_METHOD

METHOD ALARMCLEARFINISHED
END_METHOD

METHOD ALARMREAD
VAR_INPUT
	DIWHICHROW : DINT;
	STATICDATA : AlarmStorageStaticData;
END_VAR
END_METHOD

METHOD BEFOREREADING
VAR_INPUT
	USICOUNTLATCHVARIABLES : USINT;
END_VAR
END_METHOD

METHOD LATCHVARIABLEREAD
VAR_INPUT
	DIWHICHROW : DINT;
	USIWHICHVARIABLE : USINT;
	LILATCHVARVALUE : LINT;
	ILATCHVARTYPE : TypeClass;
	XVALUENULL : BOOL;
END_VAR
END_METHOD

METHOD READINGDATACOMPLETED
END_METHOD

METHOD GETNUMBEROFLATCHVARIABLES : USINT
END_METHOD

METHOD GETROOTPAGE : CAA.IDENT
VAR_INPUT
	EWHICHALARMSTORAGEOBJECT : EAlarmStorageObject;
END_VAR
END_METHOD

METHOD ISONLYONEALARMCLASSSELECTED : BOOL
END_METHOD

METHOD ISONLYONEALARMGROUPSELECTED : BOOL
END_METHOD

METHOD PREPAREDATABASEACCESS : STO.ERROR
END_METHOD

METHOD TBLALARMCURSORCLOSE : STO.ERROR
VAR_INPUT
	EERRORFROMPREVIOUSPROCESSING : STO.ERROR;
END_VAR
END_METHOD

METHOD TBLALARMCURSORMOVE : STO.ERROR
VAR_INPUT
	EDIRECTION : STO.DIRECTION;
END_VAR
VAR_OUTPUT
	XEOF : BOOL;
END_VAR
END_METHOD

METHOD TBLALARMCURSOROPEN : STO.ERROR
VAR_INPUT
	FILTERCRITERIA : REFERENCE TO VisuFbAlarmFilterCriteria;
END_VAR
END_METHOD

METHOD TBLALARMCURSOROPEN2 : STO.ERROR
VAR_INPUT
	IDINDEX : CAA.IDENT;
END_VAR
END_METHOD

METHOD TBLALARMCURSORSETPOSITION : STO.ERROR
VAR_INPUT
	FILTERCRITERIA : REFERENCE TO VisuFbAlarmFilterCriteria;
	BROWIDVALID : BOOL;
	DIROWID : DINT;
END_VAR
END_METHOD

METHOD TBLALARMGETLATCHVARTYPE : STO.ERROR
VAR_INPUT
	IDWHICHCOLUMN : CAA.IDENT;
	USIWHICHLATCHVAR : USINT;
END_VAR
VAR_OUTPUT
	BYTYPE : BYTE;
	XNULL : BOOL;
END_VAR
END_METHOD

METHOD TBLALARMGETLATCHVARVALUE : STO.ERROR
VAR_INPUT
	IDWHICHCOLUMN : CAA.IDENT;
	USIWHICHLATCHVAR : USINT;
END_VAR
VAR_OUTPUT
	LIVALUE : LINT;
	XNULL : BOOL;
END_VAR
END_METHOD

METHOD TBLALARMGETMINMAXROWIDS : BOOL
VAR_OUTPUT
	IDROWMIN : LINT;
	IDROWMAX : LINT;
	EERROR : STO.ERROR;
END_VAR
END_METHOD

METHOD TBLALARMGETROWCOUNT : CAA.COUNT
VAR_OUTPUT
	EERROR : STO.ERROR;
END_VAR
END_METHOD

METHOD TBLALARMGETTIMESTAMPVALUE : LINT
VAR_INPUT
	IDWHICHCOLUMN : CAA.IDENT;
END_VAR
VAR_OUTPUT
	EERROR : STO.ERROR;
END_VAR
END_METHOD

METHOD TBLALARMGET_DINT : STO.ERROR
VAR_INPUT
	IDWHICHCOLUMN : CAA.IDENT;
	IWHICHCOLUMN : INT;
END_VAR
VAR_OUTPUT
	DIVALUE : DINT;
	XNULL : BOOL;
END_VAR
END_METHOD

METHOD TBLALARMGET_LINT : STO.ERROR
VAR_INPUT
	IDWHICHCOLUMN : CAA.IDENT;
	IWHICHCOLUMN : INT;
END_VAR
VAR_OUTPUT
	LIVALUE : LINT;
	XNULL : BOOL;
END_VAR
END_METHOD

METHOD TBLALARMGET_SINT : STO.ERROR
VAR_INPUT
	IDWHICHCOLUMN : CAA.IDENT;
	IWHICHCOLUMN : INT;
END_VAR
VAR_OUTPUT
	SIVALUE : SINT;
	XNULL : BOOL;
END_VAR
END_METHOD

METHOD TBLALARMISNOTEMPTY : BOOL
VAR_OUTPUT
	EERROR : STO.ERROR;
END_VAR
END_METHOD

METHOD TBLALARMROWGETCURRENT : STO.ERROR
END_METHOD

METHOD TBLALARMROWGETCURRENTID : DINT
END_METHOD

METHOD TBLALARMROWISVALID : BOOL
END_METHOD

METHOD TBLALARMROWRELEASE : STO.ERROR
VAR_INPUT
	EERRORFROMPREVIOUSPROCESSING : STO.ERROR;
END_VAR
END_METHOD

METHOD TBLALARMROWSELECT : STO.ERROR
VAR_INPUT
	IDROW : CAA.IDENT;
	XDOERRORHANDLING : BOOL;
END_VAR
END_METHOD

METHOD TBLALARMTABLECLOSE : STO.ERROR
END_METHOD

METHOD TBLALARMTABLEISOPEN : BOOL
END_METHOD

METHOD TBLALARMTABLEOPEN : STO.ERROR
VAR_INPUT
	XREADONLY : BOOL;
END_VAR
END_METHOD

METHOD TBLLATCHVARSTRINGSCLOSEIFNEEDED : STO.ERROR
VAR_INPUT
	EERRORFROMPREVIOUSPROCESSING : STO.ERROR;
END_VAR
END_METHOD

METHOD TBLLATCHVARSTRINGSCURSORSEARCHROWID : STO.ERROR
VAR_INPUT
	LIROWID : LINT;
END_VAR
END_METHOD

METHOD TBLLATCHVARSTRINGSGET_TEXT : STO.ERROR
VAR_INPUT
	IDWHICHCOLUMN : CAA.IDENT;
	IWHICHCOLUMN : INT;
END_VAR
VAR_OUTPUT
	XNULL : BOOL;
END_VAR
VAR_IN_OUT
	TXTVALUE : STO.TEXT;
END_VAR
END_METHOD

METHOD TBLLATCHVARSTRINGSOPENIFNEEDED : STO.ERROR
END_METHOD

METHOD TBLLATCHVARSTRINGSROWGETCURRENT : STO.ERROR
END_METHOD

METHOD TBLLATCHVARSTRINGSROWRELEASE : STO.ERROR
VAR_INPUT
	EERRORFROMPREVIOUSPROCESSING : STO.ERROR;
END_VAR
END_METHOD

METHOD TEXTCOPYTOSTRING : STO.ERROR
VAR_INPUT
	XFREE : BOOL;
END_VAR
VAR_IN_OUT
	TXTVALUE : STO.TEXT;
	SVALUE : STRING(1);
	SZVALUE : CAA.SIZE;
END_VAR
END_METHOD

METHOD TEXTCOPYTOWSTRING : STO.ERROR
VAR_INPUT
	XFREE : BOOL;
END_VAR
VAR_IN_OUT
	TXTVALUE : STO.TEXT;
	WSVALUE : WSTRING(1);
	SZVALUE : CAA.SIZE;
END_VAR
END_METHOD

METHOD TRANSACTIONBEGIN : STO.ERROR
VAR_INPUT
	XREADONLY : BOOL;
END_VAR
END_METHOD

METHOD TRANSACTIONBEGINFAILED : BOOL
END_METHOD

METHOD TRANSACTIONEND
VAR_INPUT
	EERRORFROMPREVIOUSPROCESSING : STO.ERROR;
END_VAR
END_METHOD

METHOD TBLALARMGET_INT : STO.ERROR
VAR_INPUT
	IDWHICHCOLUMN : CAA.IDENT;
	IWHICHCOLUMN : INT;
END_VAR
VAR_OUTPUT
	IVALUE : INT;
	XNULL : BOOL;
END_VAR
END_METHOD

METHOD TBLVERSIONGETCURRENT : STO.ERROR
VAR_OUTPUT
	IVERSION : INT;
END_VAR
END_METHOD

METHOD GETRELEVANTFILTERDATA
VAR_OUTPUT
	EDBBYTEORDER : EAlarmByteOrder;
END_VAR
END_METHOD

METHOD TBLALARMCURSORSEARCHROWID : STO.ERROR
VAR_INPUT
	IDROW : DINT;
END_VAR
END_METHOD

METHOD TBLGETBYTEORDER : STO.ERROR
VAR_OUTPUT
	EBYTEORDER : EAlarmByteOrder;
END_VAR
END_METHOD

METHOD TBLVERSIONGETCURRENT2 : STO.ERROR
VAR_OUTPUT
	IVERSION : INT;
	EDBUSED : EDBType;
END_VAR
END_METHOD

METHOD TBLALARMGETCOMMENTVALUE : STO.ERROR
VAR_INPUT
	IDWHICHCOLUMN : CAA.IDENT;
	IWHICHCOLUMN : INT;
END_VAR
VAR_OUTPUT
	XNULL : BOOL;
END_VAR
VAR_IN_OUT
	WSVALUE : WSTRING(2000);
END_VAR
END_METHOD

METHOD GETALARMCLASSID : BOOL
VAR_INPUT
	DIINDEXALARM : DINT;
END_VAR
VAR_OUTPUT
	UDIALARMCLASSID : UDINT;
END_VAR
END_METHOD

METHOD GETALARMGROUPID : BOOL
VAR_INPUT
	DIINDEXALARM : DINT;
END_VAR
VAR_OUTPUT
	UDIALARMGROUPID : UDINT;
END_VAR
END_METHOD

METHOD GETALARMID : BOOL
VAR_INPUT
	DIINDEXALARM : DINT;
END_VAR
VAR_OUTPUT
	UDIALARMID : UDINT;
END_VAR
END_METHOD

METHOD GETLATCHVARTYPE : BOOL
VAR_INPUT
	DIINDEXALARM : DINT;
	IWHICHLATCHVARIABLE : INT;
END_VAR
VAR_OUTPUT
	BYTYPE : BYTE;
END_VAR
END_METHOD

METHOD GETLATCHVARVALUE : BOOL
VAR_INPUT
	DIINDEXALARM : DINT;
	IWHICHLATCHVARIABLE : INT;
END_VAR
VAR_OUTPUT
	LIVALUE : LINT;
END_VAR
END_METHOD

METHOD GETPRIORITY : BOOL
VAR_INPUT
	DIINDEXALARM : DINT;
END_VAR
VAR_OUTPUT
	USIPRIORITY : USINT;
END_VAR
END_METHOD

METHOD GETROWID : BOOL
VAR_INPUT
	DIINDEXALARM : DINT;
END_VAR
VAR_OUTPUT
	DIROWID : DINT;
END_VAR
END_METHOD

METHOD GETSTATE : BOOL
VAR_INPUT
	DIINDEXALARM : DINT;
END_VAR
VAR_OUTPUT
	BYSTATE : BYTE;
END_VAR
END_METHOD

METHOD GETTSACK : BOOL
VAR_INPUT
	DIINDEXALARM : DINT;
END_VAR
VAR_OUTPUT
	LITIMESTAMP : TIMESTAMP;
END_VAR
END_METHOD

METHOD GETTSACTIVE : BOOL
VAR_INPUT
	DIINDEXALARM : DINT;
END_VAR
VAR_OUTPUT
	LITIMESTAMP : TIMESTAMP;
END_VAR
END_METHOD

METHOD GETTSINACTIVE : BOOL
VAR_INPUT
	DIINDEXALARM : DINT;
END_VAR
VAR_OUTPUT
	LITIMESTAMP : TIMESTAMP;
END_VAR
END_METHOD

METHOD GETTSLAST : BOOL
VAR_INPUT
	DIINDEXALARM : DINT;
END_VAR
VAR_OUTPUT
	LITIMESTAMP : TIMESTAMP;
END_VAR
END_METHOD

METHOD GETTRIGGERVALUE : BOOL
VAR_INPUT
	DIINDEXALARM : DINT;
END_VAR
VAR_OUTPUT
	LIVALUE : LINT;
END_VAR
END_METHOD

METHOD GETTRIGGERVALUETYPE : BOOL
VAR_INPUT
	DIINDEXALARM : DINT;
END_VAR
VAR_OUTPUT
	BYTYPE : BYTE;
END_VAR
END_METHOD

METHOD GETREMOTEDEVICENAME : BOOL
VAR_INPUT
	DIINDEXALARM : DINT;
END_VAR
VAR_OUTPUT
	SNAME : STRING(255);
END_VAR
END_METHOD

METHOD GETCOMMENT : BOOL
VAR_INPUT
	DIINDEXALARM : DINT;
END_VAR
VAR_OUTPUT
	WSCOMMENT : WSTRING(255);
END_VAR
END_METHOD

METHOD GETUSERID : BOOL
VAR_INPUT
	DIINDEXALARM : DINT;
END_VAR
VAR_OUTPUT
	WSUSERID : WSTRING(255);
END_VAR
END_METHOD

METHOD TRYGETALARMPTRBYROWID : BOOL
VAR_INPUT
	IDROW : CAA.IDENT;
END_VAR
VAR_OUTPUT
	PALICURRALARM : POINTER TO ARRAY [0..0] OF LINT;
END_VAR
END_METHOD

METHOD WILLEXCEEDLIMIT : BOOL
END_METHOD

METHOD PRVAPPLYCIRCULARBUFFERMAPPING : DINT
VAR_INPUT
	DICURSORINDEX : DINT;
END_VAR
END_METHOD

METHOD PRVCOMPUTEBUFFERSIZE : UDINT
VAR_INPUT
	UDICOUNTALARMS : UDINT;
	USICOUNTLATCHVARIABLES : USINT;
END_VAR
VAR_OUTPUT
	UDICOUNTROWSTOALLOC : UDINT;
END_VAR
END_METHOD

METHOD PRVENLARGEBUFFERIFNECCESARY
END_METHOD

METHOD PRVFREEALLCOMMENT
VAR_INPUT
	PALICURRALARM : POINTER TO ARRAY [0..0] OF LINT;
END_VAR
END_METHOD

METHOD PRVFREECOMMENT : BOOL
VAR_INPUT
	PPWFREE : POINTER TO POINTER TO WSTRING;
END_VAR
END_METHOD

METHOD PRVGETLATCHVARTYPEOFFSET : UDINT
VAR_INPUT
	IWHICHLATCHVARIABLE : INT;
END_VAR
END_METHOD

METHOD PRVGETLATCHVARVALUEOFFSET : UDINT
VAR_INPUT
	IWHICHLATCHVARIABLE : INT;
END_VAR
END_METHOD

METHOD PRVGETTIMESTAMP : BOOL
VAR_INPUT
	DIINDEXALARM : DINT;
	UDITIMESTAMPOFFSET : UDINT;
END_VAR
VAR_OUTPUT
	LITIMESTAMP : TIMESTAMP;
END_VAR
END_METHOD

METHOD PRVPARTITION : DINT
VAR_INPUT
	DILEFT : DINT;
	DIRIGHT : DINT;
	ITFCOMPARER : IAlarmStorageDataComparer;
END_VAR
END_METHOD

METHOD PRVQUICKSORT
VAR_INPUT
	DIFIRST : DINT;
	DILAST : DINT;
	ITFCOMPARER : IAlarmStorageDataComparer;
END_VAR
END_METHOD

METHOD PRVSEARCHROWID : BOOL
VAR_INPUT
	DIROWID : DINT;
END_VAR
VAR_OUTPUT
	DIINDEX : DINT;
END_VAR
END_METHOD

METHOD PRVSORTALARMS
END_METHOD

METHOD PRVALLOC : POINTER TO DWORD
VAR_INPUT
	UDISIZE : UDINT;
	PUDIRESULT : POINTER TO RTS_IEC_RESULT;
END_VAR
END_METHOD

METHOD PRVDISPLAYSIZE
END_METHOD

METHOD PRVFREE : BOOL
VAR_INPUT
	PBLOCK : POINTER TO DWORD;
END_VAR
END_METHOD

METHOD PRVSETALARMID
VAR_INPUT
	UDIALARMID : UDINT;
END_VAR
END_METHOD

METHOD PRVSETCLASSID
VAR_INPUT
	UDIALARMCLASSID : UDINT;
END_VAR
END_METHOD

METHOD PRVSETCOMMENTVALUE
VAR_INPUT
	PWSCMT : POINTER TO WSTRING;
	OFFSET : UDINT;
END_VAR
END_METHOD

METHOD PRVSETGROUPID
VAR_INPUT
	UDIALARMGROUPID : UDINT;
END_VAR
END_METHOD

METHOD PRVSETLATCHVARTYPE
VAR_INPUT
	IWHICHLATCHVARIABLE : INT;
	ITYPE : TypeClass;
	XVALUENULL : BOOL;
END_VAR
END_METHOD

METHOD PRVSETLATCHVARVALUE
VAR_INPUT
	IWHICHLATCHVARIABLE : INT;
	LIVALUE : LINT;
END_VAR
END_METHOD

METHOD PRVSETLATCHVARVALUES
VAR_INPUT
	ALARM : AlarmStorageRow;
	XADD : BOOL;
END_VAR
END_METHOD

METHOD PRVSETOFFSETACK
VAR_INPUT
	IOFFSET : INT;
END_VAR
END_METHOD

METHOD PRVSETOFFSETACTIVE
VAR_INPUT
	IOFFSET : INT;
END_VAR
END_METHOD

METHOD PRVSETOFFSETINACTIVE
VAR_INPUT
	IOFFSET : INT;
END_VAR
END_METHOD

METHOD PRVSETOFFSETLAST
VAR_INPUT
	IOFFSET : INT;
END_VAR
END_METHOD

METHOD PRVSETPRIORITY
VAR_INPUT
	USIPRIORITY : USINT;
END_VAR
END_METHOD

METHOD PRVSETREMOTEDEVICE
VAR_INPUT
	LIVALUE : LINT;
END_VAR
END_METHOD

METHOD PRVSETROWID
VAR_INPUT
	DWROWID : DWORD;
END_VAR
END_METHOD

METHOD PRVSETSTATE
VAR_INPUT
	BYSTATE : BYTE;
END_VAR
END_METHOD

METHOD PRVSETTSACK
VAR_INPUT
	LITIMESTAMP : TIMESTAMP;
END_VAR
END_METHOD

METHOD PRVSETTSACTIVE
VAR_INPUT
	LITIMESTAMP : TIMESTAMP;
END_VAR
END_METHOD

METHOD PRVSETTSINACTIVE
VAR_INPUT
	LITIMESTAMP : TIMESTAMP;
END_VAR
END_METHOD

METHOD PRVSETTSLAST
VAR_INPUT
	LITIMESTAMP : TIMESTAMP;
END_VAR
END_METHOD

METHOD PRVSETTRIGGERVALUE
VAR_INPUT
	LIVALUE : LINT;
END_VAR
END_METHOD

METHOD PRVSETTRIGGERVALUETYPE
VAR_INPUT
	ITYPE : TypeClass;
END_VAR
END_METHOD

(* ---- ALARMSTORAGEMANAGER.fb ---- *)
FUNCTION_BLOCK ALARMSTORAGEMANAGER
VAR
	M_ALARMSTORAGE : STI.Storage;
	M_ITFSTORAGE : STO.IStorage;
	M_ITFTABLE : STO.ITable;
	M_ADWROOTPAGES : ARRAY [EAlarmStorageObject.IX_MIN..EAlarmStorageObject.IX_LAST] OF CAA.IDENT;
	M_XROOTPAGESDETERMINED : BOOL;
	M_UDICOUNTLATCHVARIABLES : CAA.COUNT;
	WRITEACCESSNECESSARY : BOOL;
END_VAR
END_FUNCTION_BLOCK

METHOD BEGINTRANSACTION : STO.ITransaction
VAR_INPUT
	XREADONLY : BOOL;
END_VAR
VAR_OUTPUT
	EERROR : STO.ERROR;
END_VAR
END_METHOD

METHOD CLOSETABLE
VAR_INPUT
	ITFTABLE : STO.ITable;
END_VAR
END_METHOD

METHOD ENDTRANSACTION
VAR_INPUT
	ITFTRANSACTION : STO.ITransaction;
	EERROR : STO.ERROR;
END_VAR
END_METHOD

METHOD FB_EXIT : BOOL
VAR_INPUT
	BINCOPYCODE : BOOL;
END_VAR
END_METHOD

METHOD GETCOLUMNIDENTIFIER : CAA.IDENT
VAR_INPUT
	IDCOLUMN : CAA.IDENT;
END_VAR
END_METHOD

METHOD GETNUMBEROFLATCHVARIABLES : CAA.COUNT
VAR_INPUT
	IDBVERSION : INT;
	UDICOUNTCOLUMNSTBLALARM : CAA.COUNT;
END_VAR
END_METHOD

METHOD GETSTORAGE : STO.IStorage
END_METHOD

METHOD OPENTABLE : STO.ITable
VAR_INPUT
	XREADONLY : BOOL;
END_VAR
VAR_OUTPUT
	EERROR : STO.ERROR;
END_VAR
END_METHOD

METHOD DETERMINEROOTPAGES : STO.ERROR
END_METHOD

METHOD GETROOTPAGE : CAA.IDENT
VAR_INPUT
	EDATABASEOBJECT : EAlarmStorageObject;
END_VAR
END_METHOD

METHOD ISREADY : BOOL
END_METHOD

METHOD RESET
END_METHOD

METHOD CLOSESTORAGE
END_METHOD

METHOD DETERMINEROOTPAGESOPENSTORAGE : STO.ERROR
VAR_OUTPUT
	XREOPENREADONLY : BOOL;
END_VAR
END_METHOD

METHOD PRVCHECKJOURNAL
END_METHOD

METHOD PRVHELPGETDATABASEFILEPATH : CAA.FILENAME
END_METHOD

METHOD PRVOPENSTORAGE : STO.ERROR
VAR_INPUT
	XREADONLY : BOOL;
END_VAR
END_METHOD

METHOD PROTCLOSECURSOR : STO.ERROR
VAR_INPUT
	EERRORFROMPREVIOUSPROCESSING : STO.ERROR;
	ICALLINGMETHOD : INT;
END_VAR
VAR_IN_OUT
	ITFCURSOR : STO.ICursor;
END_VAR
END_METHOD

METHOD PROTGETEXCLUSIVETRANSACTION : STO.ITransaction
VAR_INPUT
	ICOUNTRETRIES : INT;
END_VAR
VAR_OUTPUT
	EERROR : STO.ERROR;
END_VAR
END_METHOD

METHOD PROTRELEASEROW : STO.ERROR
VAR_INPUT
	EERRORFROMPREVIOUSPROCESSING : STO.ERROR;
	ICALLINGMETHOD : INT;
END_VAR
VAR_IN_OUT
	ITFROW : STO.IRow;
END_VAR
END_METHOD

(* ---- ALARMSTORAGEQUEUE.fb ---- *)
FUNCTION_BLOCK ALARMSTORAGEQUEUE
VAR
	_PAQUEUE : POINTER TO ARRAY [0..0] OF AlarmStorageRow;
	_IQUEUESIZE : UDINT;
	_INEWESTPOS : UDINT := 0;
	_IOLDESTPOS : UDINT := 0;
	_IITEMCOUNT : UDINT := 0;
	_ALARMSTORAGEROWPROVIDER : AlarmStorageRowProvider;
	_UICOUNTEVENTS : UDINT;
	_PAINITIALQUEUE : POINTER TO AlarmStorageRow;
	_XKEEPOLDVALUES : BOOL;
	_XFIXQUEUENECESSARY : BOOL;
	COUNTALARMSTOINSERT : UDINT;
	COUNTEVENTSTOINSERT : UDINT;
END_VAR
END_FUNCTION_BLOCK

METHOD CANPOSTALARM : BOOL
END_METHOD

METHOD CLEAR
END_METHOD

METHOD FB_EXIT : BOOL
VAR_INPUT
	BINCOPYCODE : BOOL;
END_VAR
END_METHOD

METHOD FB_INIT : BOOL
VAR_INPUT
	BINITRETAINS : BOOL;
	BINCOPYCODE : BOOL;
END_VAR
END_METHOD

METHOD FIXAFTERONLINECHANGEIFNECESSARY
VAR_INPUT
	STORAGE : IDatabaseFileAlarmStorage;
END_VAR
END_METHOD

METHOD GETCURRENTALARM : AlarmStorageRow
END_METHOD

METHOD INIT
VAR_INPUT
	PQUEUEDATA : POINTER TO AlarmStorageRow;
	NUMQUEUEENTRIES : UDINT;
END_VAR
END_METHOD

METHOD ISEMPTY : BOOL
END_METHOD

METHOD ONLINECHANGEDONE
END_METHOD

METHOD ONLINECHANGEPREPARE
END_METHOD

METHOD POSTALARM : BOOL
VAR_INPUT
	ITFALARM : IAlarm;
	ITFDATABASEFILEALARMSTORAGE : IDatabaseFileAlarmStorage;
	ESTATE : AlarmState;
	EPREVSTATE : AlarmState;
	XFORCEUPDATE : BOOL;
END_VAR
VAR_OUTPUT
	ROW : AlarmStorageRow;
END_VAR
END_METHOD

METHOD REMOVECURRENTALARM
END_METHOD

METHOD TRYTOENLARGEQUEUE
END_METHOD

METHOD ASSIGNINITVALUES
END_METHOD

METHOD RESETSTOREDREFERENCES
END_METHOD

METHOD TRYTOENLARGEQUEUEHELP
VAR_INPUT
	KEEPNEWESTPOS : BOOL;
END_VAR
END_METHOD

METHOD PRVGETTYPEDVALUE
VAR_INPUT
	ITFTYPEDVALUE : ITypedValue;
END_VAR
VAR_OUTPUT
	BYTYPECLASS : BYTE;
	LIVALUE : LINT;
END_VAR
END_METHOD

(* ---- ALARMSTORAGEREADER.fb ---- *)
FUNCTION_BLOCK ALARMSTORAGEREADER EXTENDS AlarmStorageManager
VAR_INPUT
	_HLOCK : RTS_IEC_HANDLE := RTS_INVALID_HANDLE;
END_VAR
VAR
	M_DATABASEACCESS : SQLiteDatabaseAccess;
	M_ROWIDITERATOR : AlarmStorageReaderRowIdIterator;
	M_ITFALARMSTORAGEREADERCONSUMER : IAlarmStorageReaderConsumer;
	M_ITFALARMSTORAGEMANAGER : IAlarmStorageManager := THIS^;
	M_EBYTEORDER : EAlarmByteOrder := EAlarmByteOrder.Unknown;
	M_ALATCHVARIABLES : ARRAY [1..2] OF LatchVariable;
	M_AWSLATCHVARVALUE : ARRAY [0..1] OF WSTRING(255);
	M_PALATCHVARSTRINGALLOC : POINTER TO ARRAY [0..10] OF WSTRING(255);
	M_PALATCHVARALLOC : POINTER TO ARRAY [0..10] OF LatchVariable;
	M_ICOUNTLATCHVARALLOC : INT;
	M_LOCKRESULT : RTS_IEC_RESULT;
	M_SWHOHASLOCK : STRING;
END_VAR
END_FUNCTION_BLOCK

METHOD ADDALARMSTORAGELISTENER : EAlarmStorageReaderErrors
VAR_INPUT
	ITFALARMSTORAGELISTENER : IAlarmStorageListener;
END_VAR
END_METHOD

METHOD CONTINUEREADING : EAlarmStorageReaderErrors
VAR_INPUT
	LITIMSTAMPFROM : LINT;
	LITIMSTAMPTO : LINT;
	XREADASCENDING : BOOL;
	ITFALARMSTORAGEREADERCONSUMER : IAlarmStorageReaderConsumer;
END_VAR
END_METHOD

METHOD FB_EXIT : BOOL
VAR_INPUT
	BINCOPYCODE : BOOL;
END_VAR
END_METHOD

METHOD FB_INIT : BOOL
VAR_INPUT
	BINITRETAINS : BOOL;
	BINCOPYCODE : BOOL;
END_VAR
END_METHOD

METHOD GETALARMSFROMSTORAGE : STO.ERROR
VAR_INPUT
	ISKIPROWS : INT;
	IMAXROWS : INT;
	FILTERCRITERIA : REFERENCE TO VisuFbAlarmFilterCriteria;
	ITFALARMDATABLOCK : IAlarmDataBlockBase2;
END_VAR
VAR_IN_OUT
	BROWIDVALID : BOOL;
	DIROWID : DINT;
END_VAR
END_METHOD

METHOD GETALARMSFROMSTORAGE2 : STO.ERROR
VAR_INPUT
	ITFDATABASEACCESS : IDatabaseAccess;
	ISKIPROWS : INT;
	IMAXROWS : INT;
	FILTERCRITERIA : REFERENCE TO VisuFbAlarmFilterCriteria;
	ITFALARMDATABLOCK : IAlarmDataBlockBase2;
END_VAR
VAR_IN_OUT
	BROWIDVALID : BOOL;
	DIROWID : DINT;
END_VAR
END_METHOD

METHOD GETALARMSFROMSTORAGE3 : STO.ERROR
VAR_INPUT
	ITFDATABASEACCESS : IDatabaseAccess3;
	DWROWIDLATEST : DWORD;
	IMAXROWS : INT;
	ITFALARMTRAVERSALCONSUMER : IAlarmTraversalConsumer;
END_VAR
END_METHOD

METHOD GETALARMSFROMSTORAGE4 : STO.ERROR
VAR_INPUT
	ITFDATABASEACCESS : IDatabaseAccess3;
	ITFALARMTRAVERSALCONSUMER : IAlarmTraversalConsumer;
END_VAR
END_METHOD

METHOD GETALARMSFROMSTORAGE5 : STO.ERROR
VAR_INPUT
	DISKIPROWS : DINT;
	DIMAXROWS : DINT;
	FILTERCRITERIA : REFERENCE TO VisuFbAlarmFilterCriteria;
	ITFALARMDATABLOCK : IAlarmDataBlockBase2;
END_VAR
VAR_IN_OUT
	BROWIDVALID : BOOL;
	DIROWID : DINT;
END_VAR
END_METHOD

METHOD GETALARMSFROMSTORAGE6 : STO.ERROR
VAR_INPUT
	ITFDATABASEACCESS : IDatabaseAccess;
	DISKIPROWS : DINT;
	DIMAXROWS : DINT;
	FILTERCRITERIA : REFERENCE TO VisuFbAlarmFilterCriteria;
	ITFALARMDATABLOCK : IAlarmDataBlockBase2;
END_VAR
VAR_IN_OUT
	BROWIDVALID : BOOL;
	DIROWID : DINT;
END_VAR
END_METHOD

METHOD GETCOUNTALARMSFROMSTORAGE : DINT
VAR_INPUT
	FILTERCRITERIA : REFERENCE TO VisuFbAlarmFilterCriteria;
	ITFALARMDATABLOCK : IAlarmDataBlockBase2;
END_VAR
VAR_OUTPUT
	EERROR : STO.ERROR;
	DWCOUNTLATCHVARIABLESINSTORAGE : CAA.COUNT;
END_VAR
END_METHOD

METHOD GETCOUNTALLALARMSFROMSTORAGE : CAA.COUNT
VAR_OUTPUT
	EERROR : STO.ERROR;
END_VAR
END_METHOD

METHOD GETFIRSTLASTROWID : EAlarmStorageReaderErrors
VAR_OUTPUT
	DIROWIDFIRST : DINT;
	DIROWIDLAST : DINT;
END_VAR
END_METHOD

METHOD GETMINMAXTIMESTAMPS : EAlarmStorageReaderErrors
VAR_OUTPUT
	LIMINTIMESTAMP : LINT;
	LIMAXTIMESTAMP : LINT;
	XTABLEISEMPTY : BOOL;
	UDICOUNTALARMS : UDINT;
END_VAR
END_METHOD

METHOD READ : EAlarmStorageReaderErrors
VAR_INPUT
	LITIMSTAMPFROM : LINT;
	LITIMSTAMPTO : LINT;
	XREADASCENDING : BOOL;
	ITFALARMSTORAGEREADERCONSUMER : IAlarmStorageReaderConsumer;
END_VAR
END_METHOD

METHOD REMOVEALARMSTORAGELISTENER : EAlarmStorageReaderErrors
VAR_INPUT
	ITFALARMSTORAGELISTENER : IAlarmStorageListener;
END_VAR
END_METHOD

METHOD SEMAPHOREACQUIRE
VAR_INPUT
	SWHO : STRING;
END_VAR
END_METHOD

METHOD SEMAPHORERELEASE
VAR_INPUT
	SWHO : STRING;
END_VAR
END_METHOD

METHOD PRVALLOCLATCHVARS
VAR_INPUT
	ICNTVAR : INT;
END_VAR
END_METHOD

METHOD PRVDOCONTINUEREADING : BOOL
VAR_INPUT
	DIROWCOUNTER : DINT;
END_VAR
END_METHOD

METHOD PRVFINDROWID : CAA.IDENT
VAR_INPUT
	ITFDATABASEACCESS : IDatabaseAccess;
	XSEARCHFIRST : BOOL;
END_VAR
VAR_OUTPUT
	EERROR : STO.ERROR;
END_VAR
END_METHOD

METHOD PRVFREELATCHVARS
END_METHOD

METHOD PRVREAD : EAlarmStorageReaderErrors
VAR_INPUT
	LITIMSTAMPFROM : LINT;
	LITIMSTAMPTO : LINT;
	XREADASCENDING : BOOL;
END_VAR
END_METHOD

METHOD PRVREADALARMCOMMENT
VAR_INPUT
	IDWHICHCOLUMN : CAA.IDENT;
	ITFDATABASEACCESS4 : IDatabaseAccess4;
END_VAR
VAR_IN_OUT
	EERROR : STO.ERROR;
	CMTBUFFER : AlarmComment;
END_VAR
END_METHOD

METHOD PRVREADLATCHVARSTRING2 : STO.ERROR
VAR_INPUT
	LIROWID : LINT;
	ITFDATABASEACCESS : IDatabaseAccess;
	BYLATCHVARTYPE : BYTE;
	PBVARVALUE : POINTER TO BYTE;
	ISZVARVALUE : INT;
END_VAR
END_METHOD

METHOD PRVREADLATCHVARSTRING : STO.ERROR
VAR_INPUT
	LIROWID : LINT;
	ITFDATABASEACCESS : IDatabaseAccess;
	BYLATCHVARTYPE : BYTE;
END_VAR
VAR_OUTPUT
	CBPSTRING : CharBufferPtr;
END_VAR
END_METHOD

METHOD PRVRETRIEVELATCHVARVALUE : STO.ERROR
VAR_INPUT
	ITFDATABASEACCESS : IDatabaseAccess;
	ITFALARMMETAOBJECTSTUB3 : IAlarmMetaObjectStub3;
	USIWHICHLATCHVAR : USINT;
END_VAR
END_METHOD

METHOD PRVTBLALARMFINDTIMESTAMP : STO.ERROR
VAR_INPUT
	ITFDATABASEACCESS : IDatabaseAccess;
	LITIMSTAMP : LINT;
	XUSENEXTROW : BOOL;
END_VAR
VAR_OUTPUT
	IDROWTIMSTAMP : CAA.IDENT;
END_VAR
END_METHOD

(* ---- ALARMSTORAGEREADERROWIDITERATOR.fb ---- *)
FUNCTION_BLOCK ALARMSTORAGEREADERROWIDITERATOR
VAR
	M_IDROWTBLALARMFROM : CAA.IDENT;
	M_IDROWTBLALARMTO : CAA.IDENT;
	M_IDROWCURR : CAA.IDENT;
	M_XITERATEASCENDING : BOOL;
	M_IDLASTPROCESSEDROWID : CAA.IDENT := AlarmConstants.INVALID_ROWID;
	M_LITIMESTAMP : LINT;
END_VAR
END_FUNCTION_BLOCK

METHOD GETNEXTROWID : CAA.IDENT
END_METHOD

METHOD GETSAVEDSTATE : LINT
END_METHOD

METHOD HASNEXTROWID : BOOL
END_METHOD

METHOD HASSAVEDSTATE : BOOL
END_METHOD

METHOD INITIALIZE
VAR_INPUT
	IDROWTBLALARMFROM : CAA.IDENT;
	IDROWTBLALARMTO : CAA.IDENT;
	XITERATEASCENDING : BOOL;
END_VAR
END_METHOD

METHOD SAVESTATE
VAR_INPUT
	IDLASTPROCESSEDROWID : CAA.IDENT;
	LITIMESTAMP : LINT;
END_VAR
END_METHOD

(* ---- ALARMSTORAGEROW.fb ---- *)
FUNCTION_BLOCK ALARMSTORAGEROW
VAR_INPUT
	UDIALARMID : UDINT;
	UDIALARMCLASSID : UDINT;
	UDIALARMGROUPID : UDINT;
	LITIMESTAPLAST : TIMESTAMP;
	LITIMESTAPACTIVE : TIMESTAMP;
	LITIMESTAPINACTIVE : TIMESTAMP;
	LITIMESTAPACKNOWLEDGE : TIMESTAMP;
	IOFFSETLAST : INT := -1;
	IOFFSETACTIVE : INT := -1;
	IOFFSETINACTIVE : INT := -1;
	IOFFSETACKNOWLEDGE : INT := -1;
	USIPRIORITY : USINT;
	ESTATE : AlarmState;
	EPREVSTATE : AlarmState;
	BYTRIGGERVALUETYPE : BYTE;
	LITRIGGERVALUEVAL : LINT;
	PLATCHVARIABLES : POINTER TO ARRAY [0..10] OF LatchVariable;
	USICOUNTLATCHVARIABLES : USINT;
	ITFALARM : IAlarm;
	ITFDATABASEFILEALARMSTORAGE : IDatabaseFileAlarmStorage;
	IDROW : CAA.IDENT;
	XIDROWVALID : BOOL;
	XFORCEUPDATE : BOOL;
	SREMOTEDEVICENAME : STRING;
	CMTACTIVE : AlarmComment;
	CMTACTIVEACK : AlarmComment;
	CMTWAITINGCONF : AlarmComment;
	CMTNORMAL : AlarmComment;
	XINVALID : BOOL;
END_VAR
END_FUNCTION_BLOCK

METHOD DERIVEALARMREFERENCE
END_METHOD

METHOD GETLATCHVARVALUE
VAR_INPUT
	USIWHICHLATCHVAR : USINT;
END_VAR
VAR_OUTPUT
	BYTYPE : BYTE;
	LIVALUE : LINT;
END_VAR
END_METHOD

METHOD RESETALARMCOMMENTS : BOOL
END_METHOD

METHOD SETLATCHVARVALUE
VAR_INPUT
	USIWHICHLATCHVAR : USINT;
	BYTYPE : BYTE;
	LIVALUE : LINT;
END_VAR
END_METHOD

(* ---- ALARMSTORAGEROWPROVIDER.fb ---- *)
FUNCTION_BLOCK ALARMSTORAGEROWPROVIDER
VAR
	M_PAALARMSTORAGEROWS : POINTER TO ARRAY [0..100] OF AlarmStorageRow;
	M_ICOUNTROWS : UDINT;
	M_PALATCHVARIABLES : POINTER TO ARRAY [0..100] OF LatchVariable;
	M_ICOUNTLATCHVARIABLES : UDINT;
	COMPONENT : STRING := 'AlarmStorageRowProvider';
END_VAR
END_FUNCTION_BLOCK

METHOD ALLOCATEALARMSTORAGEROWARRAY : BOOL
VAR_INPUT
	IREQUIREDARRAYSIZE : UDINT;
	USICOUNTLATCHVARIABLES : USINT;
	PACURRENTQUEUE : POINTER TO AlarmStorageRow;
	ICURRENTQUEUESIZE : UDINT;
	ICURRENTREADINDEX : UDINT;
END_VAR
VAR_OUTPUT
	PANEWQUEUE : POINTER TO ARRAY [0..0] OF AlarmStorageRow;
	INEWQUEUESIZE : UDINT;
END_VAR
END_METHOD

METHOD COPYQUEUECONTENT : BOOL
VAR_INPUT
	PACURRENTQUEUE : POINTER TO AlarmStorageRow;
	ICURRENTQUEUESIZE : UDINT;
	ICURRENTREADINDEX : UDINT;
	PANEWALARMSTORAGEROWS : POINTER TO AlarmStorageRow;
	INEWQUEUESIZE : UDINT;
	PANEWLATCHVARIABLES : POINTER TO LatchVariable;
	USICOUNTLATCHVARIABLES : USINT;
END_VAR
END_METHOD

METHOD FB_EXIT : BOOL
VAR_INPUT
	BINCOPYCODE : BOOL;
END_VAR
END_METHOD

METHOD FREEBUFFER
VAR_INPUT
	PPBYBUFFER : POINTER TO POINTER TO BYTE;
	PICOUNT : POINTER TO INT;
END_VAR
END_METHOD

METHOD FREEBUFFERS
END_METHOD

(* ---- ALLOCATOR.fb ---- *)
FUNCTION_BLOCK ALLOCATOR
VAR_INPUT
	SCOMPONENT : STRING;
END_VAR
VAR
	DITOTMEM : DINT;
	TOTMEM : DINT;
END_VAR
END_FUNCTION_BLOCK

METHOD ALLOCANDCOPYWSTRING : POINTER TO WSTRING
VAR_INPUT
	PWSWHO : POINTER TO WSTRING;
END_VAR
END_METHOD

METHOD ALLOCBYTES : POINTER TO BYTE
VAR_INPUT
	UXISIZE : __UXINT;
	SWHO : STRING;
END_VAR
END_METHOD

METHOD ALLOCPROXYFBALARMCONTAINER : POINTER TO AlarmContainer
VAR_INPUT
	SWHO : STRING;
END_VAR
END_METHOD

METHOD ALLOCPROXYFBALARMMETAOBJECTSTUB : POINTER TO ProxyFbAlarmMetaObjectStub
VAR_INPUT
	SWHO : STRING;
END_VAR
END_METHOD

METHOD ALLOCPROXYSTRUCTALARMCLASSDESCRIPTION : POINTER TO ProxyStructAlarmClass
VAR_INPUT
	SWHO : STRING;
END_VAR
END_METHOD

METHOD ALLOCPROXYSTRUCTALARMDESCRIPTION : POINTER TO ProxyStructAlarm
VAR_INPUT
	SWHO : STRING;
END_VAR
END_METHOD

METHOD ALLOCPROXYSTRUCTALARMGROUPDESCRIPTION : POINTER TO ProxyStructAlarmGroup
VAR_INPUT
	SWHO : STRING;
END_VAR
END_METHOD

METHOD ALLOCPROXYSTRUCTHISTORICALALARMACTIVE : POINTER TO ProxyStructHistoricalAlarmActive
VAR_INPUT
	SWHO : STRING;
END_VAR
END_METHOD

METHOD ALLOCVALUETYPEBUNDLE : POINTER TO ValueTypeBundle
VAR_INPUT
	SWHO : STRING;
END_VAR
END_METHOD

METHOD FREEBYTES
VAR_INPUT
	PTR : POINTER TO BYTE;
	UXISIZE : __UXINT;
END_VAR
END_METHOD

METHOD FREEPROXYFBALARMCONTAINER
VAR_INPUT
	PREQ : POINTER TO AlarmContainer;
END_VAR
END_METHOD

METHOD FREEPROXYFBALARMMETAOBJECTSTUB
VAR_INPUT
	PREQ : POINTER TO ProxyFbAlarmMetaObjectStub;
END_VAR
END_METHOD

METHOD FREEPROXYSTRUCTALARMCLASSDESCRIPTION
VAR_INPUT
	PREQ : POINTER TO ProxyStructAlarmGroup;
END_VAR
END_METHOD

METHOD FREEPROXYSTRUCTALARMDESCRIPTION
VAR_INPUT
	PREQ : POINTER TO ProxyStructAlarm;
END_VAR
END_METHOD

METHOD FREEPROXYSTRUCTALARMGROUPDESCRIPTION
VAR_INPUT
	PREQ : POINTER TO ProxyStructAlarmClass;
END_VAR
END_METHOD

METHOD FREEPROXYSTRUCTHISTORICALALARMACTIVE
VAR_INPUT
	PREQ : POINTER TO ProxyStructHistoricalAlarmActive;
END_VAR
END_METHOD

METHOD FREEVALUETYPEBUNDLE
VAR_INPUT
	PREQ : POINTER TO ValueTypeBundle;
END_VAR
END_METHOD

(* ---- BINTAGWRITERALARMMETAOBJECTSTUB.fb ---- *)
FUNCTION_BLOCK BINTAGWRITERALARMMETAOBJECTSTUB
VAR
	M_ITFTAGGEDSERVICEWRITER : ITaggedServiceWriter;
	M_LITIMESTAMPACKNOWLEDGE : Timestamp;
	M_LITIMESTAMPACTIVE : Timestamp;
	M_LITIMESTAMPINACTIVE : Timestamp;
	M_LITIMESTAMPLAST : Timestamp;
	M_ITFTYPEDVALUETRIGGER : ITypedValue;
	M_IOFFSETACKNOWLEDGE : INT := -1;
	M_IOFFSETACTIVE : INT := -1;
	M_IOFFSETINACTIVE : INT := -1;
	M_IOFFSETLAST : INT := -1;
	M_PALATCHVARIABLES : POINTER TO ARRAY [0..0] OF LatchVariable;
	M_ICOUNTLATCHVARIABLES : INT;
	M_ISTATE : INT;
	M_UDIALARMID : UDINT;
	M_UDIALARMGROUPID : UDINT;
	OFFSETACKNOWLEDGE : INT;
	OFFSETACTIVE : INT;
	OFFSETINACTIVE : INT;
	OFFSETLAST : INT;
END_VAR
END_FUNCTION_BLOCK

METHOD INITIALIZE
VAR_INPUT
	ITFTAGGEDSERVICEWRITER : ITaggedServiceWriter;
END_VAR
END_METHOD

METHOD SETLATCHVARIABLESBUFFER
VAR_INPUT
	PALATCHVARIABLES : POINTER TO ARRAY [0..0] OF LatchVariable;
	ICOUNTLATCHVARIABLES : INT;
END_VAR
END_METHOD

METHOD SETLATCHVAR1VALUE
VAR_INPUT
	ITFTYPEDVALUELATCHVAR1 : ITypedValue;
END_VAR
END_METHOD

METHOD SETLATCHVAR2VALUE
VAR_INPUT
	ITFTYPEDVALUELATCHVAR2 : ITypedValue;
END_VAR
END_METHOD

METHOD SETSTATE
VAR_INPUT
	ISTATE : INT;
END_VAR
END_METHOD

METHOD SETTIMESTAMPACKNOWLEDGE
VAR_INPUT
	LITIMESTAMPACKNOWLEDGE : Timestamp;
END_VAR
END_METHOD

METHOD SETTIMESTAMPACTIVE
VAR_INPUT
	LITIMESTAMPACTIVE : Timestamp;
END_VAR
END_METHOD

METHOD SETTIMESTAMPINACTIVE
VAR_INPUT
	LITIMESTAMPINACTIVE : Timestamp;
END_VAR
END_METHOD

METHOD SETTIMESTAMPLAST
VAR_INPUT
	LITIMESTAMPLAST : Timestamp;
END_VAR
END_METHOD

METHOD SETTRIGGERVALUE
VAR_INPUT
	ITFTYPEDVALUETRIGGER : ITypedValue;
END_VAR
END_METHOD

METHOD GETCOUNTLATCHVARIABLES : USINT
END_METHOD

METHOD GETLATCHVARVALUE : ITypedValue2
VAR_INPUT
	IWHICHLATCHVAR : INT;
END_VAR
END_METHOD

METHOD SETLATCHVARVALUE
VAR_INPUT
	IWHICHLATCHVAR : INT;
	ITFTYPEDVALUELATCHVAR : ITypedValue;
END_VAR
END_METHOD

METHOD SETALARM
VAR_INPUT
	PALARM : POINTER TO Alarm;
END_VAR
END_METHOD

METHOD FILLINGCOMPLETED : UDINT
END_METHOD

METHOD PRVGETTYPE : BYTE
VAR_INPUT
	ITFTYPEDVALUE : ITypedValue;
END_VAR
END_METHOD

METHOD PRVGETVALUE : LWORD
VAR_INPUT
	ITFTYPEDVALUE : ITypedValue;
END_VAR
END_METHOD

METHOD PRVWRITELATCHVARIABLE
VAR_INPUT
	IWHICHLATCHVAR : INT;
END_VAR
END_METHOD

METHOD GETALARMGROUP : STRING
END_METHOD

METHOD GETCHECKSUM : UDINT
END_METHOD

METHOD GETCURRENTVALUE : ITypedValue
END_METHOD

METHOD GETID : ALARM_ID
END_METHOD

METHOD GETLATCHVAR1VALUE : ITypedValue
END_METHOD

METHOD GETLATCHVAR2VALUE : ITypedValue
END_METHOD

METHOD GETSTATE : INT
END_METHOD

METHOD GETTIMESTAMPACKNOWLEDGE : Timestamp
END_METHOD

METHOD GETTIMESTAMPACTIVE : Timestamp
END_METHOD

METHOD GETTIMESTAMPINACTIVE : Timestamp
END_METHOD

METHOD GETTIMESTAMPLAST : Timestamp
END_METHOD

METHOD GETTRIGGERVALUE : ITypedValue
END_METHOD

METHOD SETACKNOWLEDGE
VAR_INPUT
	BACKNOWLEDGEMULTIPLE : BOOL;
END_VAR
END_METHOD

METHOD SETALARMGROUP
VAR_INPUT
	SALARMGROUP : STRING;
END_VAR
END_METHOD

METHOD SETCURRENTLREALVALUE
VAR_INPUT
	LRVALUE : LREAL;
END_VAR
END_METHOD

METHOD SETID
VAR_INPUT
	UIID : ALARM_ID;
END_VAR
END_METHOD

METHOD SWAPVALUES
END_METHOD

METHOD GETALARM : POINTER TO Alarm
END_METHOD

METHOD SETCURRENTVALUE
VAR_INPUT
	ITFTYPEDVALUECURRENT : ITypedValue;
END_VAR
END_METHOD

(* ---- BINTAGWRITERDATABLOCK.fb ---- *)
FUNCTION_BLOCK BINTAGWRITERDATABLOCK
VAR
	M_BINTAGWRITERALARMMETAOBJECTSTUB : BinTagWriterAlarmMetaObjectStub;
	M_ICOUNTROWS : INT;
END_VAR
END_FUNCTION_BLOCK

METHOD GETALARMMETAOBJECTSTUB : IAlarmMetaObjectStub3
VAR_INPUT
	IROW : INT;
	IOFFSET : INT;
END_VAR
END_METHOD

METHOD GETCOUNTROWS : INT
END_METHOD

METHOD INITIALIZE
VAR_INPUT
	ITFTAGGEDSERVICEWRITER : ITaggedServiceWriter;
END_VAR
END_METHOD

METHOD SETCOUNTROWS : BOOL
VAR_INPUT
	ICOUNT : INT;
END_VAR
END_METHOD

METHOD SETLATCHVARIABLESBUFFER
VAR_INPUT
	PALATCHVARIABLES : POINTER TO ARRAY [0..0] OF LatchVariable;
	ICOUNTLATCHVARIABLES : INT;
END_VAR
END_METHOD

METHOD HASALARMS : BOOL
END_METHOD

METHOD SETTOTALCOUNTROWS : BOOL
VAR_INPUT
	DICOUNT : DINT;
END_VAR
END_METHOD

(* ---- CHANGEOBSERVATIONTYPE.fb ---- *)
FUNCTION_BLOCK CHANGEOBSERVATIONTYPE
VAR_INPUT
	M_UIID : ALARM_ID;
	M_ITFCHANGEEVALUATOR : IChangeEvaluator;
END_VAR
END_FUNCTION_BLOCK

METHOD ISACTIVE : BOOL
VAR_INPUT
	ECURRSTATE : AlarmState;
END_VAR
END_METHOD

METHOD ISIMMEDIATELYACTIVE : BOOL
END_METHOD

(* ---- COMMENTCOMPARER.fb ---- *)
FUNCTION_BLOCK COMMENTCOMPARER EXTENDS TSLastComparer
END_FUNCTION_BLOCK

METHOD COMPARE : INT
VAR_INPUT
	DIINDEXALARM1 : DINT;
	DIINDEXALARM2 : DINT;
END_VAR
END_METHOD

(* ---- COMPONENTREGISTRATOR.fb ---- *)
FUNCTION_BLOCK COMPONENTREGISTRATOR
VAR
	_HCOMPONENT : RTS_IEC_HANDLE;
	CMINVALIDHANDLE : RTS_IEC_HANDLE := 16#FFFFFFFF;
END_VAR
END_FUNCTION_BLOCK

METHOD FB_EXIT : BOOL
VAR_INPUT
	BINCOPYCODE : BOOL;
END_VAR
END_METHOD

METHOD FB_INIT
VAR_INPUT
	BINITRETAINS : BOOL;
	BINCOPYCODE : BOOL;
END_VAR
END_METHOD

(* ---- CONVERTIECTYPEDLITERAL.fb ---- *)
FUNCTION_BLOCK CONVERTIECTYPEDLITERAL
VAR
	CH_PLUS : BYTE := 16#2B;
	CH_MINUS : BYTE := 16#2D;
	CH_POINT : BYTE := 16#2E;
	CH_0 : BYTE := 16#30;
	CH_1 : BYTE := 16#31;
	CH_2 : BYTE := 16#32;
	CH_3 : BYTE := 16#33;
	CH_4 : BYTE := 16#34;
	CH_5 : BYTE := 16#35;
	CH_6 : BYTE := 16#36;
	CH_7 : BYTE := 16#37;
	CH_8 : BYTE := 16#38;
	CH_9 : BYTE := 16#39;
	CH_COLON : BYTE := 16#3A;
	CH_A : BYTE := 16#41;
	CH_B : BYTE := 16#42;
	CH_C : BYTE := 16#43;
	CH_D : BYTE := 16#44;
	CH_E : BYTE := 16#45;
	CH_F : BYTE := 16#46;
	CH_H : BYTE := 16#48;
	CH_M : BYTE := 16#4D;
	CH_N : BYTE := 16#4E;
	CH_S : BYTE := 16#53;
	CH_U : BYTE := 16#55;
END_VAR
END_FUNCTION_BLOCK

METHOD CONVERT : INT
VAR_INPUT
	SLITERAL : STRING(255);
	XCONVERTCHECK : BOOL;
END_VAR
VAR_OUTPUT
	VTYPE : Visu_Types;
	LIVALUE : LINT;
	RVALUE : REAL;
	LRVALUE : LREAL;
END_VAR
END_METHOD

METHOD TEST : STRING
END_METHOD

METHOD CONVERTOLD : INT
VAR_INPUT
	PLITERAL : POINTER TO STRING(255);
END_VAR
VAR_OUTPUT
	VTYPE : Visu_Types;
	LIVALUE : LINT;
	RVALUE : REAL;
	LRVALUE : LREAL;
END_VAR
END_METHOD

METHOD PRVANALYSEDURATIONVALUE : LINT
VAR_INPUT
	PNUMBER : POINTER TO STRING(255);
	LIUNIT : LINT;
END_VAR
END_METHOD

METHOD PRVGETDATE : BOOL
VAR_INPUT
	PTOKEN : POINTER TO STRING(255);
END_VAR
VAR_OUTPUT
	LIDATE : LINT;
END_VAR
END_METHOD

METHOD PRVGETDATEANDTIME : BOOL
VAR_INPUT
	PTOKEN : POINTER TO STRING(255);
END_VAR
VAR_OUTPUT
	LIDT : LINT;
END_VAR
END_METHOD

METHOD PRVGETDURATION : BOOL
VAR_INPUT
	PTOKEN : POINTER TO STRING(255);
END_VAR
VAR_OUTPUT
	LIDURATION : LINT;
END_VAR
END_METHOD

METHOD PRVGETFACTOR
VAR_INPUT
	LIBASE : LINT;
	PSUB : POINTER TO STRING;
END_VAR
VAR_OUTPUT
	LIFACTOR : LINT;
END_VAR
END_METHOD

METHOD PRVGETLREAL : BOOL
VAR_INPUT
	PTOKEN : POINTER TO STRING(255);
END_VAR
VAR_OUTPUT
	LRVALUE : LREAL;
END_VAR
END_METHOD

METHOD PRVGETNUMERICAL : BOOL
VAR_INPUT
	PTOKEN : POINTER TO STRING(255);
	XSIGNALLOWED : BOOL;
END_VAR
VAR_OUTPUT
	LIVALUE : LINT;
	SBASE16VALUE : STRING;
END_VAR
END_METHOD

METHOD PRVGETREAL : BOOL
VAR_INPUT
	PTOKEN : POINTER TO STRING(255);
END_VAR
VAR_OUTPUT
	RVALUE : REAL;
END_VAR
END_METHOD

METHOD PRVGETTIMEOFDAY : BOOL
VAR_INPUT
	PTOKEN : POINTER TO STRING(255);
END_VAR
VAR_OUTPUT
	LITOD : LINT;
END_VAR
END_METHOD

METHOD PRVINTTODATE : BOOL
VAR_INPUT
	IDAY : INT;
	IMONTH : INT;
	IYEAR : INT;
END_VAR
VAR_OUTPUT
	UIDAYS : UINT;
END_VAR
END_METHOD

METHOD PRVSPLIT
VAR_INPUT
	PSTRING : POINTER TO STRING(255);
	SSPLITCHAR : STRING;
END_VAR
VAR_OUTPUT
	SLEFT : STRING(255);
	SRIGHT : STRING(255);
END_VAR
END_METHOD

(* ---- DATABASEACCESSERRORHANDLER.fb ---- *)
FUNCTION_BLOCK DATABASEACCESSERRORHANDLER
VAR_INPUT
	M_UIDISKFULLDATABASEACCESSSUSPENDTIME : UINT;
END_VAR
VAR
	M_XLOGERRORS : BOOL := TRUE;
	M_XDATABASEACCESSENABLED : BOOL := TRUE;
	M_DWTIMESTAMPFIRSTDISKFULLEVENT : DWORD;
END_VAR
END_FUNCTION_BLOCK

METHOD ERRORHANDLING
VAR_INPUT
	IFUNCTION : INT;
	IERRCODE : INT;
END_VAR
END_METHOD

METHOD ISDATABASEACCESSENABLED : BOOL
END_METHOD

METHOD ISSEARCHNOTFOUNDERROR : BOOL
VAR_INPUT
	EERROR : STO.ERROR;
END_VAR
END_METHOD

METHOD SQLITEERRORHANDLING
VAR_INPUT
	IFUNCTION : INT;
	EERROR : STO.ERROR;
	IACTION : INT;
END_VAR
END_METHOD

METHOD SQLITEERRORHANDLINGSEARCHING
VAR_INPUT
	IFUNCTION : INT;
	EERROR : STO.ERROR;
	IACTION : INT;
END_VAR
END_METHOD

METHOD PRVGETFUNCTIONNAME : STRING
VAR_INPUT
	IFUNCTION : INT;
END_VAR
END_METHOD
